FUNCTION "ROLL_PB2" : Void
{ S7_Optimized_Access := 'TRUE' }
VERSION : 0.1
VAR_TEMP
    r : Bool;
    a1 : Word;
    a2 : Word;
    activeDataBlock : Int;
    comparisonResults : Array[0..0] of Bool;
END_VAR
BEGIN
    #r := FALSE;
    #a1 := W#16#0000;
    #a2 := W#16#0000;
    #activeDataBlock := 0;
    // PB2, STEP 5 network 1
    #r := ((NOT "ROLL_State".M[0, 1]) AND "ROLL_State".S5Timers[11].Q);
    "ROLL_State".M[4, 1] := #r;
    // PB2, STEP 5 network 2
    #r := ((NOT "ROLL_State".M[4, 1]) OR "ROLL_IO".Input[1, 0]);
    "ROLL_State".M[3, 1] := #r;
    // PB2, STEP 5 network 3
    #r := ((((NOT "ROLL_State".M[31, 4]) AND "ROLL_IO".Input[0, 4] AND "ROLL_State".M[4, 1]) OR "ROLL_State".M[31, 5]) AND "ROLL_IO".Input[0, 2]);
    "ROLL_State".M[4, 4] := #r;
    // PB2, STEP 5 network 4
    #r := (NOT "ROLL_IO".Input[11, 7]);
    IF #r THEN "ROLL_State".M[5, 0] := TRUE; END_IF;
    #r := "ROLL_State".M[3, 1];
    IF #r THEN "ROLL_State".M[5, 0] := FALSE; END_IF;
    // PB2, STEP 5 network 5
    #r := (NOT "ROLL_IO".Input[13, 5]);
    IF #r THEN "ROLL_State".M[5, 1] := TRUE; END_IF;
    #r := "ROLL_State".M[3, 1];
    IF #r THEN "ROLL_State".M[5, 1] := FALSE; END_IF;
    // PB2, STEP 5 network 6
    #r := (NOT "ROLL_IO".Input[13, 0]);
    IF #r THEN "ROLL_State".M[5, 2] := TRUE; END_IF;
    #r := "ROLL_State".M[3, 1];
    IF #r THEN "ROLL_State".M[5, 2] := FALSE; END_IF;
    // PB2, STEP 5 network 7
    #r := (NOT "ROLL_IO".Input[8, 5]);
    IF #r THEN "ROLL_State".M[5, 3] := TRUE; END_IF;
    #r := "ROLL_State".M[3, 1];
    IF #r THEN "ROLL_State".M[5, 3] := FALSE; END_IF;
    // PB2, STEP 5 network 8
    #r := "ROLL_State".M[0, 3];
    IF #r THEN "ROLL_State".M[5, 4] := TRUE; END_IF;
    #r := "ROLL_State".M[3, 1];
    IF #r THEN "ROLL_State".M[5, 4] := FALSE; END_IF;
    // PB2, STEP 5 network 9
    #r := "ROLL_State".M[0, 3];
    IF #r THEN "ROLL_State".M[5, 5] := TRUE; END_IF;
    #r := "ROLL_State".M[3, 1];
    IF #r THEN "ROLL_State".M[5, 5] := FALSE; END_IF;
    // PB2, STEP 5 network 10
    #r := "ROLL_IO".Input[3, 6];
    IF #r THEN "ROLL_State".M[5, 6] := TRUE; END_IF;
    #r := "ROLL_State".M[3, 1];
    IF #r THEN "ROLL_State".M[5, 6] := FALSE; END_IF;
    // PB2, STEP 5 network 11
    #r := (NOT "ROLL_IO".Input[3, 7]);
    IF #r THEN "ROLL_State".M[5, 7] := TRUE; END_IF;
    #r := "ROLL_State".M[3, 1];
    IF #r THEN "ROLL_State".M[5, 7] := FALSE; END_IF;
    // PB2, STEP 5 network 12
    #r := (NOT "ROLL_IO".Input[5, 2]);
    IF #r THEN "ROLL_State".M[6, 0] := TRUE; END_IF;
    #r := ("ROLL_IO".Input[5, 2] AND "ROLL_State".M[3, 1]);
    IF #r THEN "ROLL_State".M[6, 0] := FALSE; END_IF;
    // PB2, STEP 5 network 13
    #r := ((NOT "ROLL_IO".Input[5, 3]) AND "ROLL_State".S5Timers[31].Q);
    IF #r THEN "ROLL_State".M[6, 1] := TRUE; END_IF;
    #r := "ROLL_State".M[3, 1];
    IF #r THEN "ROLL_State".M[6, 1] := FALSE; END_IF;
    // PB2, STEP 5 network 14
    #r := (NOT "ROLL_IO".Input[5, 4]);
    IF #r THEN "ROLL_State".M[6, 2] := TRUE; END_IF;
    #r := ("ROLL_IO".Input[5, 4] AND "ROLL_State".M[3, 1]);
    IF #r THEN "ROLL_State".M[6, 2] := FALSE; END_IF;
    // PB2, STEP 5 network 15
    #r := ((NOT "ROLL_IO".Input[5, 5]) AND "ROLL_State".M[40, 5] AND "ROLL_State".S5Timers[17].Q);
    IF #r THEN "ROLL_State".M[6, 3] := TRUE; END_IF;
    #r := "ROLL_State".M[3, 1];
    IF #r THEN "ROLL_State".M[6, 3] := FALSE; END_IF;
    // PB2, STEP 5 network 16
    #r := ((NOT "ROLL_IO".Input[6, 0]) AND "ROLL_State".S5Timers[32].Q);
    IF #r THEN "ROLL_State".M[6, 4] := TRUE; END_IF;
    #r := "ROLL_State".M[3, 1];
    IF #r THEN "ROLL_State".M[6, 4] := FALSE; END_IF;
    // PB2, STEP 5 network 17
    #r := ((NOT "ROLL_IO".Input[6, 2]) AND "ROLL_State".S5Timers[33].Q);
    IF #r THEN "ROLL_State".M[6, 5] := TRUE; END_IF;
    #r := "ROLL_State".M[3, 1];
    IF #r THEN "ROLL_State".M[6, 5] := FALSE; END_IF;
    // PB2, STEP 5 network 18
    #r := "ROLL_State".M[0, 3];
    IF #r THEN "ROLL_State".M[6, 6] := TRUE; END_IF;
    #r := "ROLL_State".M[3, 1];
    IF #r THEN "ROLL_State".M[6, 6] := FALSE; END_IF;
    // PB2, STEP 5 network 19
    #r := ((NOT "ROLL_State".M[0, 3]) AND "ROLL_State".S5Timers[35].Q);
    IF #r THEN "ROLL_State".M[6, 7] := TRUE; END_IF;
    #r := "ROLL_State".M[3, 1];
    IF #r THEN "ROLL_State".M[6, 7] := FALSE; END_IF;
    // PB2, STEP 5 network 20
    #r := ((NOT "ROLL_State".M[0, 3]) AND "ROLL_State".S5Timers[36].Q);
    IF #r THEN "ROLL_State".M[7, 0] := TRUE; END_IF;
    #r := "ROLL_State".M[3, 1];
    IF #r THEN "ROLL_State".M[7, 0] := FALSE; END_IF;
    // PB2, STEP 5 network 21
    #r := ((NOT "ROLL_State".M[0, 3]) AND "ROLL_State".M[48, 1] AND "ROLL_State".S5Timers[37].Q);
    IF #r THEN "ROLL_State".M[7, 1] := TRUE; END_IF;
    #r := "ROLL_State".M[3, 1];
    IF #r THEN "ROLL_State".M[7, 1] := FALSE; END_IF;
    // PB2, STEP 5 network 22
    #r := ((NOT "ROLL_State".M[0, 3]) AND "ROLL_State".S5Timers[38].Q);
    IF #r THEN "ROLL_State".M[7, 2] := TRUE; END_IF;
    #r := "ROLL_State".M[3, 1];
    IF #r THEN "ROLL_State".M[7, 2] := FALSE; END_IF;
    // PB2, STEP 5 network 23
    #r := ((NOT "ROLL_IO".Input[5, 6]) AND "ROLL_State".S5Timers[16].Q);
    IF #r THEN "ROLL_State".M[7, 3] := TRUE; END_IF;
    #r := ("ROLL_IO".Input[5, 6] AND "ROLL_State".M[3, 1]);
    IF #r THEN "ROLL_State".M[7, 3] := FALSE; END_IF;
    // PB2, STEP 5 network 24
    #r := "ROLL_State".M[0, 3];
    IF #r THEN "ROLL_State".M[7, 4] := TRUE; END_IF;
    #r := "ROLL_State".M[3, 1];
    IF #r THEN "ROLL_State".M[7, 4] := FALSE; END_IF;
    // PB2, STEP 5 network 25
    #r := "ROLL_State".M[0, 3];
    IF #r THEN "ROLL_State".M[7, 5] := TRUE; END_IF;
    #r := "ROLL_State".M[3, 1];
    IF #r THEN "ROLL_State".M[7, 5] := FALSE; END_IF;
    // PB2, STEP 5 network 26
    #r := "ROLL_State".M[0, 3];
    IF #r THEN "ROLL_State".M[7, 6] := TRUE; END_IF;
    #r := "ROLL_State".M[3, 1];
    IF #r THEN "ROLL_State".M[7, 6] := FALSE; END_IF;
    // PB2, STEP 5 network 27
    #r := (NOT "ROLL_IO".Input[6, 7]);
    IF #r THEN "ROLL_State".M[7, 7] := TRUE; END_IF;
    #r := "ROLL_State".M[3, 1];
    IF #r THEN "ROLL_State".M[7, 7] := FALSE; END_IF;
    // PB2, STEP 5 network 28
    #a2 := #a1;
    #a1 := W#16#1050;
    #r := ((NOT "ROLL_IO".Input[7, 6]) AND "ROLL_IO".Output[20, 5]);
    "ROLL_TimerOp"(Number := 30, Operation := 0, Signal := #r, Preset := #a1);
    #r := "ROLL_State".S5Timers[30].Q;
    IF #r THEN "ROLL_State".M[8, 6] := TRUE; END_IF;
    #r := "ROLL_State".M[3, 1];
    IF #r THEN "ROLL_State".M[8, 6] := FALSE; END_IF;
    // PB2, STEP 5 network 29
    #r := "ROLL_State".M[0, 3];
    IF #r THEN "ROLL_State".M[8, 7] := TRUE; END_IF;
    #r := "ROLL_State".M[3, 1];
    IF #r THEN "ROLL_State".M[8, 7] := FALSE; END_IF;
    // PB2, STEP 5 network 30
    #r := ((NOT "ROLL_IO".Input[13, 7]) AND "ROLL_State".M[4, 1]);
    IF #r THEN "ROLL_State".M[9, 0] := TRUE; END_IF;
    #r := ("ROLL_IO".Input[13, 7] AND "ROLL_State".M[3, 1]);
    IF #r THEN "ROLL_State".M[9, 0] := FALSE; END_IF;
    // PB2, STEP 5 network 31
    #r := "ROLL_State".M[0, 3];
    IF #r THEN "ROLL_State".M[9, 1] := TRUE; END_IF;
    #r := "ROLL_State".M[3, 1];
    IF #r THEN "ROLL_State".M[9, 1] := FALSE; END_IF;
    // PB2, STEP 5 network 32
    #r := ((NOT "ROLL_State".M[28, 4]) AND (NOT "ROLL_State".M[31, 5]) AND (((NOT "ROLL_State".M[20, 2]) AND ("ROLL_IO".Input[123, 5] OR "ROLL_IO".Input[123, 6])) OR "ROLL_State".M[70, 2] OR "ROLL_State".M[70, 3]) AND "ROLL_IO".Input[0, 4] AND "ROLL_State".M[4, 1]);
    IF #r THEN "ROLL_State".M[9, 2] := TRUE; END_IF;
    #r := "ROLL_State".M[3, 1];
    IF #r THEN "ROLL_State".M[9, 2] := FALSE; END_IF;
    // PB2, STEP 5 network 33
    #r := ("ROLL_State".M[4, 1] AND "ROLL_State".S5Timers[19].Q);
    IF #r THEN "ROLL_State".M[9, 3] := TRUE; END_IF;
    #r := "ROLL_State".M[3, 1];
    IF #r THEN "ROLL_State".M[9, 3] := FALSE; END_IF;
    // PB2, STEP 5 network 34
    #r := (((("ROLL_State".M[20, 4] OR "ROLL_State".M[20, 5]) AND "ROLL_IO".Input[0, 1] AND "ROLL_State".M[190, 6]) OR "ROLL_State".M[31, 5]) AND "ROLL_State".S5Timers[95].Q);
    "ROLL_State".M[9, 4] := #r;
    // PB2, STEP 5 network 35
    #r := "ROLL_State".M[0, 3];
    IF #r THEN "ROLL_State".M[9, 5] := TRUE; END_IF;
    #r := "ROLL_State".M[3, 1];
    IF #r THEN "ROLL_State".M[9, 5] := FALSE; END_IF;
    // PB2, STEP 5 network 36
    #r := "ROLL_State".M[0, 3];
    IF #r THEN "ROLL_State".M[9, 6] := TRUE; END_IF;
    #r := "ROLL_State".M[3, 1];
    IF #r THEN "ROLL_State".M[9, 6] := FALSE; END_IF;
    // PB2, STEP 5 network 37
    #r := "ROLL_State".M[0, 3];
    IF #r THEN "ROLL_State".M[9, 7] := TRUE; END_IF;
    #r := "ROLL_State".M[3, 1];
    IF #r THEN "ROLL_State".M[9, 7] := FALSE; END_IF;
    // PB2, STEP 5 network 38
    #r := ((NOT "ROLL_IO".Input[12, 0]) AND "ROLL_State".M[4, 1]);
    IF #r THEN "ROLL_State".M[10, 0] := TRUE; END_IF;
    #r := (((((NOT "ROLL_State".S5Timers[11].Q) AND "ROLL_IO".Input[3, 0]) OR "ROLL_IO".Input[12, 5]) AND "ROLL_State".M[3, 1]) OR (NOT "ROLL_State".M[4, 1]) OR "ROLL_State".M[0, 7]);
    IF #r THEN "ROLL_State".M[10, 0] := FALSE; END_IF;
    // PB2, STEP 5 network 39
    #r := ((NOT "ROLL_IO".Input[12, 6]) AND "ROLL_State".M[4, 1]);
    IF #r THEN "ROLL_State".M[10, 1] := TRUE; END_IF;
    #r := (((((NOT "ROLL_State".S5Timers[11].Q) AND "ROLL_IO".Input[3, 0]) OR "ROLL_IO".Input[12, 1]) AND "ROLL_State".M[3, 1]) OR (NOT "ROLL_State".M[4, 1]) OR "ROLL_State".M[0, 7]);
    IF #r THEN "ROLL_State".M[10, 1] := FALSE; END_IF;
    // PB2, STEP 5 network 40
    #r := "ROLL_State".M[0, 3];
    IF #r THEN "ROLL_State".M[10, 2] := TRUE; END_IF;
    #r := "ROLL_State".M[3, 1];
    IF #r THEN "ROLL_State".M[10, 2] := FALSE; END_IF;
    // PB2, STEP 5 network 41
    #r := "ROLL_State".M[0, 3];
    IF #r THEN "ROLL_State".M[10, 3] := TRUE; END_IF;
    #r := "ROLL_State".M[3, 1];
    IF #r THEN "ROLL_State".M[10, 3] := FALSE; END_IF;
    // PB2, STEP 5 network 42
    #r := "ROLL_State".M[0, 3];
    IF #r THEN "ROLL_State".M[10, 4] := TRUE; END_IF;
    #r := "ROLL_State".M[3, 1];
    IF #r THEN "ROLL_State".M[10, 4] := FALSE; END_IF;
    // PB2, STEP 5 network 43
    #r := "ROLL_State".M[0, 3];
    IF #r THEN "ROLL_State".M[10, 5] := TRUE; END_IF;
    #r := "ROLL_State".M[3, 1];
    IF #r THEN "ROLL_State".M[10, 5] := FALSE; END_IF;
    // PB2, STEP 5 network 44
    #r := "ROLL_State".M[0, 3];
    IF #r THEN "ROLL_State".M[10, 6] := TRUE; END_IF;
    #r := "ROLL_State".M[3, 1];
    IF #r THEN "ROLL_State".M[10, 6] := FALSE; END_IF;
    // PB2, STEP 5 network 45
    #r := "ROLL_State".M[0, 3];
    IF #r THEN "ROLL_State".M[10, 7] := TRUE; END_IF;
    #r := "ROLL_State".M[3, 1];
    IF #r THEN "ROLL_State".M[10, 7] := FALSE; END_IF;
    // PB2, STEP 5 network 46
    #r := ("ROLL_State".M[4, 1] AND "ROLL_State".M[63, 2]);
    IF #r THEN "ROLL_State".M[11, 0] := TRUE; END_IF;
    #r := "ROLL_State".M[3, 1];
    IF #r THEN "ROLL_State".M[11, 0] := FALSE; END_IF;
    // PB2, STEP 5 network 47
    #r := ("ROLL_IO".Input[13, 3] AND "ROLL_State".M[4, 1] AND "ROLL_State".S5Timers[112].Q);
    IF #r THEN "ROLL_State".M[11, 1] := TRUE; END_IF;
    #r := "ROLL_State".M[3, 1];
    IF #r THEN "ROLL_State".M[11, 1] := FALSE; END_IF;
    // PB2, STEP 5 network 48
    #r := ((NOT "ROLL_IO".Input[13, 3]) AND "ROLL_State".M[4, 1] AND "ROLL_State".S5Timers[15].Q);
    IF #r THEN "ROLL_State".M[11, 2] := TRUE; END_IF;
    #r := "ROLL_State".M[3, 1];
    IF #r THEN "ROLL_State".M[11, 2] := FALSE; END_IF;
    // PB2, STEP 5 network 49
    #r := ("ROLL_State".M[4, 1] AND "ROLL_State".M[63, 3]);
    IF #r THEN "ROLL_State".M[11, 3] := TRUE; END_IF;
    #r := "ROLL_State".M[3, 1];
    IF #r THEN "ROLL_State".M[11, 3] := FALSE; END_IF;
    // PB2, STEP 5 network 50
    #r := ("ROLL_State".M[190, 6] AND "ROLL_State".M[23, 2] AND "ROLL_State".M[60, 3]);
    IF #r THEN "ROLL_State".M[11, 4] := TRUE; END_IF;
    #r := "ROLL_State".M[3, 1];
    IF #r THEN "ROLL_State".M[11, 4] := FALSE; END_IF;
    // PB2, STEP 5 network 51
    #r := "ROLL_State".M[0, 3];
    IF #r THEN "ROLL_State".M[11, 5] := TRUE; END_IF;
    #r := "ROLL_State".M[3, 1];
    IF #r THEN "ROLL_State".M[11, 5] := FALSE; END_IF;
    // PB2, STEP 5 network 52
    #r := "ROLL_State".M[0, 3];
    IF #r THEN "ROLL_State".M[11, 6] := TRUE; END_IF;
    #r := "ROLL_State".M[3, 1];
    IF #r THEN "ROLL_State".M[11, 6] := FALSE; END_IF;
    // PB2, STEP 5 network 53
    #r := "ROLL_State".M[0, 3];
    IF #r THEN "ROLL_State".M[11, 7] := TRUE; END_IF;
    #r := "ROLL_State".M[3, 1];
    IF #r THEN "ROLL_State".M[11, 7] := FALSE; END_IF;
    // PB2, STEP 5 network 54
    #r := (NOT "ROLL_IO".Input[8, 3]);
    IF #r THEN "ROLL_State".M[12, 0] := TRUE; END_IF;
    #r := "ROLL_State".M[3, 1];
    IF #r THEN "ROLL_State".M[12, 0] := FALSE; END_IF;
    // PB2, STEP 5 network 55
    #r := ((NOT "ROLL_IO".Input[0, 7]) AND (NOT "ROLL_IO".Input[1, 4]) AND "ROLL_State".M[4, 4]);
    IF #r THEN "ROLL_State".M[12, 1] := TRUE; END_IF;
    #r := "ROLL_State".M[3, 1];
    IF #r THEN "ROLL_State".M[12, 1] := FALSE; END_IF;
    // PB2, STEP 5 network 56
    #r := "ROLL_State".M[0, 3];
    IF #r THEN "ROLL_State".M[12, 2] := TRUE; END_IF;
    #r := "ROLL_State".M[3, 1];
    IF #r THEN "ROLL_State".M[12, 2] := FALSE; END_IF;
    // PB2, STEP 5 network 57
    #r := "ROLL_State".M[0, 3];
    IF #r THEN "ROLL_State".M[12, 3] := TRUE; END_IF;
    #r := "ROLL_State".M[3, 1];
    IF #r THEN "ROLL_State".M[12, 3] := FALSE; END_IF;
    // PB2, STEP 5 network 58
    #r := "ROLL_State".M[0, 3];
    IF #r THEN "ROLL_State".M[13, 0] := TRUE; END_IF;
    #r := "ROLL_State".M[3, 1];
    IF #r THEN "ROLL_State".M[13, 0] := FALSE; END_IF;
    // PB2, STEP 5 network 59
    #r := (NOT "ROLL_IO".Input[3, 2]);
    IF #r THEN "ROLL_State".M[13, 1] := TRUE; END_IF;
    #r := "ROLL_State".M[3, 1];
    IF #r THEN "ROLL_State".M[13, 1] := FALSE; END_IF;
    // PB2, STEP 5 network 60
    #r := ((NOT "ROLL_IO".Input[4, 7]) AND "ROLL_IO".Input[0, 1] AND "ROLL_State".M[190, 6] AND "ROLL_State".M[27, 4]);
    IF #r THEN "ROLL_State".M[13, 2] := TRUE; END_IF;
    #r := "ROLL_State".M[3, 1];
    IF #r THEN "ROLL_State".M[13, 2] := FALSE; END_IF;
    // PB2, STEP 5 network 61
    #r := (NOT "ROLL_IO".Input[5, 0]);
    IF #r THEN "ROLL_State".M[13, 3] := TRUE; END_IF;
    #r := ("ROLL_IO".Input[5, 0] AND "ROLL_State".M[3, 1]);
    IF #r THEN "ROLL_State".M[13, 3] := FALSE; END_IF;
    // PB2, STEP 5 network 62
    #r := (NOT "ROLL_IO".Input[10, 7]);
    IF #r THEN "ROLL_State".M[13, 4] := TRUE; END_IF;
    #r := ("ROLL_IO".Input[10, 7] AND "ROLL_State".M[3, 1]);
    IF #r THEN "ROLL_State".M[13, 4] := FALSE; END_IF;
    // PB2, STEP 5 network 63
    #r := (NOT "ROLL_IO".Input[4, 5]);
    IF #r THEN "ROLL_State".M[13, 7] := TRUE; END_IF;
    #r := "ROLL_State".M[3, 1];
    IF #r THEN "ROLL_State".M[13, 7] := FALSE; END_IF;
    // PB2, STEP 5 network 64
    #a2 := #a1;
    #a1 := W#16#2020;
    #r := (((NOT "ROLL_IO".Input[10, 0]) OR (NOT "ROLL_IO".Input[10, 1]) OR (NOT "ROLL_IO".Input[10, 2]) OR (NOT "ROLL_IO".Input[10, 3])) AND "ROLL_IO".Output[19, 1]);
    "ROLL_TimerOp"(Number := 50, Operation := 0, Signal := #r, Preset := #a1);
    // PB2, STEP 5 network 65
    #r := ((NOT "ROLL_IO".Input[10, 0]) AND "ROLL_State".S5Timers[50].Q);
    IF #r THEN "ROLL_State".M[14, 0] := TRUE; END_IF;
    #r := "ROLL_State".M[3, 1];
    IF #r THEN "ROLL_State".M[14, 0] := FALSE; END_IF;
    // PB2, STEP 5 network 66
    #r := ((NOT "ROLL_IO".Input[10, 1]) AND "ROLL_State".S5Timers[50].Q);
    IF #r THEN "ROLL_State".M[14, 1] := TRUE; END_IF;
    #r := "ROLL_State".M[3, 1];
    IF #r THEN "ROLL_State".M[14, 1] := FALSE; END_IF;
    // PB2, STEP 5 network 67
    #r := ((NOT "ROLL_IO".Input[10, 2]) AND "ROLL_State".S5Timers[50].Q);
    IF #r THEN "ROLL_State".M[14, 2] := TRUE; END_IF;
    #r := "ROLL_State".M[3, 1];
    IF #r THEN "ROLL_State".M[14, 2] := FALSE; END_IF;
    // PB2, STEP 5 network 68
    #r := ((NOT "ROLL_IO".Input[10, 3]) AND "ROLL_State".S5Timers[50].Q);
    IF #r THEN "ROLL_State".M[14, 3] := TRUE; END_IF;
    #r := "ROLL_State".M[3, 1];
    IF #r THEN "ROLL_State".M[14, 3] := FALSE; END_IF;
    // PB2, STEP 5 network 69
    #r := "ROLL_State".M[0, 3];
    IF #r THEN "ROLL_State".M[15, 2] := TRUE; END_IF;
    #r := "ROLL_State".M[3, 1];
    IF #r THEN "ROLL_State".M[15, 2] := FALSE; END_IF;
    // PB2, STEP 5 network 70
    #r := "ROLL_State".M[0, 3];
    IF #r THEN "ROLL_State".M[15, 3] := TRUE; END_IF;
    #r := "ROLL_State".M[3, 1];
    IF #r THEN "ROLL_State".M[15, 3] := FALSE; END_IF;
    // PB2, STEP 5 network 71
    #r := "ROLL_State".M[0, 3];
    IF #r THEN "ROLL_State".M[15, 4] := TRUE; END_IF;
    #r := "ROLL_State".M[3, 1];
    IF #r THEN "ROLL_State".M[15, 4] := FALSE; END_IF;
    // PB2, STEP 5 network 72
    #r := (NOT "ROLL_IO".Input[4, 0]);
    IF #r THEN "ROLL_State".M[15, 5] := TRUE; END_IF;
    #r := "ROLL_State".M[3, 1];
    IF #r THEN "ROLL_State".M[15, 5] := FALSE; END_IF;
    // PB2, STEP 5 network 73
    #r := (NOT "ROLL_IO".Input[4, 1]);
    IF #r THEN "ROLL_State".M[15, 6] := TRUE; END_IF;
    #r := "ROLL_State".M[3, 1];
    IF #r THEN "ROLL_State".M[15, 6] := FALSE; END_IF;
    // PB2, STEP 5 network 74
    #r := (NOT "ROLL_IO".Input[4, 2]);
    IF #r THEN "ROLL_State".M[15, 7] := TRUE; END_IF;
    #r := "ROLL_State".M[3, 1];
    IF #r THEN "ROLL_State".M[15, 7] := FALSE; END_IF;
    // PB2, STEP 5 network 75
    #r := "ROLL_State".M[16, 0];
    IF #r THEN "ROLL_State".M[16, 0] := TRUE; END_IF;
    #r := "ROLL_State".M[3, 1];
    IF #r THEN "ROLL_State".M[16, 0] := FALSE; END_IF;
    // PB2, STEP 5 network 76
    #r := "ROLL_State".M[16, 1];
    IF #r THEN "ROLL_State".M[16, 1] := TRUE; END_IF;
    #r := "ROLL_State".M[3, 1];
    IF #r THEN "ROLL_State".M[16, 1] := FALSE; END_IF;
    // PB2, STEP 5 network 77
    #r := "ROLL_State".M[16, 2];
    IF #r THEN "ROLL_State".M[16, 2] := TRUE; END_IF;
    #r := "ROLL_State".M[3, 1];
    IF #r THEN "ROLL_State".M[16, 2] := FALSE; END_IF;
    // PB2, STEP 5 network 78
    #r := ("ROLL_State".M[34, 1] AND "ROLL_State".M[4, 1]);
    IF #r THEN "ROLL_State".M[16, 3] := TRUE; END_IF;
    #r := "ROLL_State".M[3, 1];
    IF #r THEN "ROLL_State".M[16, 3] := FALSE; END_IF;
    // PB2, STEP 5 network 79
    #r := "ROLL_State".M[16, 4];
    IF #r THEN "ROLL_State".M[16, 4] := TRUE; END_IF;
    #r := ((NOT "ROLL_IO".Input[123, 1]) AND (NOT "ROLL_IO".Input[123, 4]) AND (NOT "ROLL_IO".Input[123, 5]) AND (NOT "ROLL_IO".Input[123, 6]) AND (NOT "ROLL_IO".Input[125, 0]) AND (NOT "ROLL_IO".Input[125, 1]) AND "ROLL_State".M[3, 1]);
    IF #r THEN "ROLL_State".M[16, 4] := FALSE; END_IF;
    // PB2, STEP 5 network 80
    #r := "ROLL_State".M[16, 5];
    IF #r THEN "ROLL_State".M[16, 5] := TRUE; END_IF;
    #r := "ROLL_State".M[3, 1];
    IF #r THEN "ROLL_State".M[16, 5] := FALSE; END_IF;
    // PB2, STEP 5 network 81
    #r := ((NOT "ROLL_IO".Input[3, 4]) AND "ROLL_State".M[4, 1]);
    IF #r THEN "ROLL_State".M[16, 6] := TRUE; END_IF;
    #r := ("ROLL_IO".Input[3, 4] AND "ROLL_State".M[3, 1]);
    IF #r THEN "ROLL_State".M[16, 6] := FALSE; END_IF;
    // PB2, STEP 5 network 82
    #r := ((NOT "ROLL_IO".Input[3, 1]) AND ((("ROLL_State".M[190, 5] OR "ROLL_State".M[190, 6]) AND "ROLL_IO".Input[0, 1]) OR "ROLL_State".M[4, 4]) AND "ROLL_State".M[4, 1]);
    IF #r THEN "ROLL_State".M[16, 7] := TRUE; END_IF;
    #r := "ROLL_State".M[3, 1];
    IF #r THEN "ROLL_State".M[16, 7] := FALSE; END_IF;
    // PB2, STEP 5 network 83
    #r := ((NOT "ROLL_IO".Input[3, 5]) AND "ROLL_State".M[4, 1]);
    IF #r THEN "ROLL_State".M[17, 0] := TRUE; END_IF;
    #r := ("ROLL_IO".Input[3, 5] AND "ROLL_State".M[3, 1]);
    IF #r THEN "ROLL_State".M[17, 0] := FALSE; END_IF;
    // PB2, STEP 5 network 84
    #r := "ROLL_State".M[0, 3];
    IF #r THEN "ROLL_State".M[17, 1] := TRUE; END_IF;
    #r := "ROLL_State".M[3, 1];
    IF #r THEN "ROLL_State".M[17, 1] := FALSE; END_IF;
    // PB2, STEP 5 network 85
    #r := "ROLL_State".M[0, 3];
    IF #r THEN "ROLL_State".M[17, 2] := TRUE; END_IF;
    #r := "ROLL_State".M[3, 1];
    IF #r THEN "ROLL_State".M[17, 2] := FALSE; END_IF;
    // PB2, STEP 5 network 86
    #r := "ROLL_State".M[0, 3];
    IF #r THEN "ROLL_State".M[17, 3] := TRUE; END_IF;
    #r := "ROLL_State".M[3, 1];
    IF #r THEN "ROLL_State".M[17, 3] := FALSE; END_IF;
    // PB2, STEP 5 network 87
    #r := "ROLL_State".M[0, 3];
    IF #r THEN "ROLL_State".M[17, 4] := TRUE; END_IF;
    #r := "ROLL_State".M[3, 1];
    IF #r THEN "ROLL_State".M[17, 4] := FALSE; END_IF;
    // PB2, STEP 5 network 88
    #r := "ROLL_State".M[0, 3];
    IF #r THEN "ROLL_State".M[17, 5] := TRUE; END_IF;
    #r := "ROLL_State".M[3, 1];
    IF #r THEN "ROLL_State".M[17, 5] := FALSE; END_IF;
    // PB2, STEP 5 network 89
    #r := "ROLL_State".M[0, 3];
    IF #r THEN "ROLL_State".M[17, 6] := TRUE; END_IF;
    #r := "ROLL_State".M[3, 1];
    IF #r THEN "ROLL_State".M[17, 6] := FALSE; END_IF;
    // PB2, STEP 5 network 90
    #r := "ROLL_State".M[0, 3];
    IF #r THEN "ROLL_State".M[17, 7] := TRUE; END_IF;
    #r := "ROLL_State".M[3, 1];
    IF #r THEN "ROLL_State".M[17, 7] := FALSE; END_IF;
    // PB2, STEP 5 network 91
    #r := "ROLL_State".M[0, 3];
    IF #r THEN "ROLL_State".M[18, 0] := TRUE; END_IF;
    #r := "ROLL_State".M[3, 1];
    IF #r THEN "ROLL_State".M[18, 0] := FALSE; END_IF;
    // PB2, STEP 5 network 92
    #r := ((NOT "ROLL_IO".Input[14, 0]) AND ((("ROLL_State".M[190, 5] OR "ROLL_State".M[190, 6]) AND ("ROLL_State".M[23, 0] OR "ROLL_State".M[23, 1] OR "ROLL_State".M[23, 2] OR "ROLL_State".M[23, 3])) OR ("ROLL_State".M[16, 3] AND "ROLL_State".M[31, 4] AND "ROLL_State".M[37, 2]) OR "ROLL_State".M[74, 0]));
    IF #r THEN "ROLL_State".M[18, 1] := TRUE; END_IF;
    #r := "ROLL_State".M[3, 1];
    IF #r THEN "ROLL_State".M[18, 1] := FALSE; END_IF;
    // PB2, STEP 5 network 93
    #r := "ROLL_State".M[0, 3];
    IF #r THEN "ROLL_State".M[18, 2] := TRUE; END_IF;
    #r := "ROLL_State".M[3, 1];
    IF #r THEN "ROLL_State".M[18, 2] := FALSE; END_IF;
    // PB2, STEP 5 network 94
    #r := "ROLL_State".M[0, 3];
    IF #r THEN "ROLL_State".M[18, 3] := TRUE; END_IF;
    #r := "ROLL_State".M[3, 1];
    IF #r THEN "ROLL_State".M[18, 3] := FALSE; END_IF;
    // PB2, STEP 5 network 95
    #r := "ROLL_State".M[0, 3];
    IF #r THEN "ROLL_State".M[18, 4] := TRUE; END_IF;
    #r := "ROLL_State".M[3, 1];
    IF #r THEN "ROLL_State".M[18, 4] := FALSE; END_IF;
    // PB2, STEP 5 network 96
    #r := "ROLL_State".M[0, 3];
    IF #r THEN "ROLL_State".M[18, 5] := TRUE; END_IF;
    #r := "ROLL_State".M[3, 1];
    IF #r THEN "ROLL_State".M[18, 5] := FALSE; END_IF;
    // PB2, STEP 5 network 97
    #r := "ROLL_State".M[0, 3];
    IF #r THEN "ROLL_State".M[18, 6] := TRUE; END_IF;
    #r := "ROLL_State".M[3, 1];
    IF #r THEN "ROLL_State".M[18, 6] := FALSE; END_IF;
    // PB2, STEP 5 network 98
    #r := "ROLL_State".M[0, 3];
    IF #r THEN "ROLL_State".M[18, 7] := TRUE; END_IF;
    #r := "ROLL_State".M[3, 1];
    IF #r THEN "ROLL_State".M[18, 7] := FALSE; END_IF;
    // PB2, STEP 5 network 99
    #r := "ROLL_State".M[0, 3];
    IF #r THEN "ROLL_State".M[19, 0] := TRUE; END_IF;
    #r := "ROLL_State".M[3, 1];
    IF #r THEN "ROLL_State".M[19, 0] := FALSE; END_IF;
    // PB2, STEP 5 network 100
    #r := "ROLL_State".M[0, 3];
    IF #r THEN "ROLL_State".M[19, 1] := TRUE; END_IF;
    #r := "ROLL_State".M[3, 1];
    IF #r THEN "ROLL_State".M[19, 1] := FALSE; END_IF;
    // PB2, STEP 5 network 101
    #r := "ROLL_State".M[0, 3];
    IF #r THEN "ROLL_State".M[19, 2] := TRUE; END_IF;
    #r := "ROLL_State".M[3, 1];
    IF #r THEN "ROLL_State".M[19, 2] := FALSE; END_IF;
    // PB2, STEP 5 network 102
    #r := "ROLL_State".M[0, 3];
    IF #r THEN "ROLL_State".M[19, 3] := TRUE; END_IF;
    #r := "ROLL_State".M[3, 1];
    IF #r THEN "ROLL_State".M[19, 3] := FALSE; END_IF;
    // PB2, STEP 5 network 103
    #r := "ROLL_State".M[0, 3];
    IF #r THEN "ROLL_State".M[19, 4] := TRUE; END_IF;
    #r := "ROLL_State".M[3, 1];
    IF #r THEN "ROLL_State".M[19, 4] := FALSE; END_IF;
    // PB2, STEP 5 network 104
    #r := "ROLL_State".M[0, 3];
    IF #r THEN "ROLL_State".M[19, 5] := TRUE; END_IF;
    #r := "ROLL_State".M[3, 1];
    IF #r THEN "ROLL_State".M[19, 5] := FALSE; END_IF;
    // PB2, STEP 5 network 105
    #r := "ROLL_State".M[0, 3];
    IF #r THEN "ROLL_State".M[19, 6] := TRUE; END_IF;
    #r := "ROLL_State".M[3, 1];
    IF #r THEN "ROLL_State".M[19, 6] := FALSE; END_IF;
    // PB2, STEP 5 network 106
    #r := "ROLL_State".M[0, 3];
    IF #r THEN "ROLL_State".M[19, 7] := TRUE; END_IF;
    #r := "ROLL_State".M[3, 1];
    IF #r THEN "ROLL_State".M[19, 7] := FALSE; END_IF;
    // PB2, STEP 5 network 107
    RETURN;
END_FUNCTION

FUNCTION "ROLL_PB3" : Void
{ S7_Optimized_Access := 'TRUE' }
VERSION : 0.1
VAR_TEMP
    r : Bool;
    a1 : Word;
    a2 : Word;
    activeDataBlock : Int;
    comparisonResults : Array[0..15] of Bool;
END_VAR
BEGIN
    #r := FALSE;
    #a1 := W#16#0000;
    #a2 := W#16#0000;
    #activeDataBlock := 0;
    // PB3, STEP 5 network 1
    #a2 := #a1;
    #a1 := "ROLL_GetM"(FirstByte := 239, Width := 8);
    #a2 := #a1;
    #a1 := W#16#0001;
    #comparisonResults[0] := (WORD_TO_INT(#a2) = WORD_TO_INT(#a1));
    #r := #comparisonResults[0];
    "ROLL_State".M[20, 1] := #r;
    // PB3, STEP 5 network 2
    #a2 := #a1;
    #a1 := "ROLL_GetM"(FirstByte := 239, Width := 8);
    #a2 := #a1;
    #a1 := W#16#0002;
    #comparisonResults[1] := (WORD_TO_INT(#a2) = WORD_TO_INT(#a1));
    #r := #comparisonResults[1];
    "ROLL_State".M[20, 2] := #r;
    // PB3, STEP 5 network 3
    #a2 := #a1;
    #a1 := "ROLL_GetM"(FirstByte := 239, Width := 8);
    #a2 := #a1;
    #a1 := W#16#0003;
    #comparisonResults[2] := (WORD_TO_INT(#a2) = WORD_TO_INT(#a1));
    #r := #comparisonResults[2];
    "ROLL_State".M[20, 3] := #r;
    // PB3, STEP 5 network 4
    #a2 := #a1;
    #a1 := "ROLL_GetM"(FirstByte := 239, Width := 8);
    #a2 := #a1;
    #a1 := W#16#0004;
    #comparisonResults[3] := (WORD_TO_INT(#a2) = WORD_TO_INT(#a1));
    #r := #comparisonResults[3];
    "ROLL_State".M[20, 4] := #r;
    // PB3, STEP 5 network 5
    #a2 := #a1;
    #a1 := "ROLL_GetM"(FirstByte := 239, Width := 8);
    #a2 := #a1;
    #a1 := W#16#0005;
    #comparisonResults[4] := (WORD_TO_INT(#a2) = WORD_TO_INT(#a1));
    #r := #comparisonResults[4];
    "ROLL_State".M[20, 5] := #r;
    // PB3, STEP 5 network 6
    #a2 := #a1;
    #a1 := "ROLL_GetM"(FirstByte := 239, Width := 8);
    #a2 := #a1;
    #a1 := W#16#0007;
    #comparisonResults[5] := (WORD_TO_INT(#a2) = WORD_TO_INT(#a1));
    #r := #comparisonResults[5];
    "ROLL_State".M[20, 7] := #r;
    // PB3, STEP 5 network 7
    #a2 := #a1;
    #a1 := "ROLL_GetM"(FirstByte := 239, Width := 8);
    #a2 := #a1;
    #a1 := W#16#000A;
    #comparisonResults[6] := (WORD_TO_INT(#a2) = WORD_TO_INT(#a1));
    #r := #comparisonResults[6];
    "ROLL_State".M[22, 0] := #r;
    // PB3, STEP 5 network 8
    #a2 := #a1;
    #a1 := "ROLL_GetM"(FirstByte := 239, Width := 8);
    #a2 := #a1;
    #a1 := W#16#000B;
    #comparisonResults[7] := (WORD_TO_INT(#a2) = WORD_TO_INT(#a1));
    #r := #comparisonResults[7];
    "ROLL_State".M[22, 1] := #r;
    // PB3, STEP 5 network 9
    #a2 := #a1;
    #a1 := "ROLL_GetM"(FirstByte := 239, Width := 8);
    #a2 := #a1;
    #a1 := W#16#000C;
    #comparisonResults[8] := (WORD_TO_INT(#a2) = WORD_TO_INT(#a1));
    #r := #comparisonResults[8];
    "ROLL_State".M[22, 2] := #r;
    // PB3, STEP 5 network 10
    #a2 := #a1;
    #a1 := "ROLL_GetM"(FirstByte := 239, Width := 8);
    #a2 := #a1;
    #a1 := W#16#000D;
    #comparisonResults[9] := (WORD_TO_INT(#a2) = WORD_TO_INT(#a1));
    #r := #comparisonResults[9];
    "ROLL_State".M[22, 3] := #r;
    // PB3, STEP 5 network 11
    #a2 := #a1;
    #a1 := "ROLL_GetM"(FirstByte := 239, Width := 8);
    #a2 := #a1;
    #a1 := W#16#000E;
    #comparisonResults[10] := (WORD_TO_INT(#a2) = WORD_TO_INT(#a1));
    #r := #comparisonResults[10];
    "ROLL_State".M[22, 4] := #r;
    // PB3, STEP 5 network 12
    #a2 := #a1;
    #a1 := "ROLL_GetM"(FirstByte := 239, Width := 8);
    #a2 := #a1;
    #a1 := W#16#000F;
    #comparisonResults[11] := (WORD_TO_INT(#a2) = WORD_TO_INT(#a1));
    #r := #comparisonResults[11];
    "ROLL_State".M[22, 5] := #r;
    // PB3, STEP 5 network 13
    #a2 := #a1;
    #a1 := "ROLL_GetM"(FirstByte := 239, Width := 8);
    #a2 := #a1;
    #a1 := W#16#0014;
    #comparisonResults[12] := (WORD_TO_INT(#a2) = WORD_TO_INT(#a1));
    #r := #comparisonResults[12];
    "ROLL_State".M[23, 0] := #r;
    // PB3, STEP 5 network 14
    #a2 := #a1;
    #a1 := "ROLL_GetM"(FirstByte := 239, Width := 8);
    #a2 := #a1;
    #a1 := W#16#0015;
    #comparisonResults[13] := (WORD_TO_INT(#a2) = WORD_TO_INT(#a1));
    #r := #comparisonResults[13];
    "ROLL_State".M[23, 1] := #r;
    // PB3, STEP 5 network 15
    #a2 := #a1;
    #a1 := "ROLL_GetM"(FirstByte := 239, Width := 8);
    #a2 := #a1;
    #a1 := W#16#0016;
    #comparisonResults[14] := (WORD_TO_INT(#a2) = WORD_TO_INT(#a1));
    #r := #comparisonResults[14];
    "ROLL_State".M[23, 2] := #r;
    // PB3, STEP 5 network 16
    #a2 := #a1;
    #a1 := "ROLL_GetM"(FirstByte := 239, Width := 8);
    #a2 := #a1;
    #a1 := W#16#0017;
    #comparisonResults[15] := (WORD_TO_INT(#a2) = WORD_TO_INT(#a1));
    #r := #comparisonResults[15];
    "ROLL_State".M[23, 3] := #r;
    // PB3, STEP 5 network 17
    RETURN;
END_FUNCTION

FUNCTION "ROLL_PB4" : Void
{ S7_Optimized_Access := 'TRUE' }
VERSION : 0.1
VAR_TEMP
    r : Bool;
    a1 : Word;
    a2 : Word;
    activeDataBlock : Int;
    comparisonResults : Array[0..24] of Bool;
END_VAR
BEGIN
    #r := FALSE;
    #a1 := W#16#0000;
    #a2 := W#16#0000;
    #activeDataBlock := 0;
    // PB4, STEP 5 network 1
    #a2 := #a1;
    #a1 := "ROLL_GetM"(FirstByte := 239, Width := 8);
    #a2 := #a1;
    #a1 := W#16#001E;
    #comparisonResults[0] := (WORD_TO_INT(#a2) = WORD_TO_INT(#a1));
    #r := #comparisonResults[0];
    "ROLL_State".M[23, 5] := #r;
    // PB4, STEP 5 network 2
    #a2 := #a1;
    #a1 := "ROLL_GetM"(FirstByte := 239, Width := 8);
    #a2 := #a1;
    #a1 := W#16#001F;
    #comparisonResults[1] := (WORD_TO_INT(#a2) = WORD_TO_INT(#a1));
    #r := #comparisonResults[1];
    "ROLL_State".M[23, 6] := #r;
    // PB4, STEP 5 network 3
    #a2 := #a1;
    #a1 := "ROLL_GetM"(FirstByte := 239, Width := 8);
    #a2 := #a1;
    #a1 := W#16#0023;
    #comparisonResults[2] := (WORD_TO_INT(#a2) = WORD_TO_INT(#a1));
    #r := #comparisonResults[2];
    "ROLL_State".M[24, 0] := #r;
    // PB4, STEP 5 network 4
    #a2 := #a1;
    #a1 := "ROLL_GetM"(FirstByte := 239, Width := 8);
    #a2 := #a1;
    #a1 := W#16#0024;
    #comparisonResults[3] := (WORD_TO_INT(#a2) = WORD_TO_INT(#a1));
    #r := #comparisonResults[3];
    "ROLL_State".M[24, 1] := #r;
    // PB4, STEP 5 network 5
    #a2 := #a1;
    #a1 := "ROLL_GetM"(FirstByte := 239, Width := 8);
    #a2 := #a1;
    #a1 := W#16#0025;
    #comparisonResults[4] := (WORD_TO_INT(#a2) = WORD_TO_INT(#a1));
    #r := #comparisonResults[4];
    "ROLL_State".M[24, 2] := #r;
    // PB4, STEP 5 network 6
    #a2 := #a1;
    #a1 := "ROLL_GetM"(FirstByte := 239, Width := 8);
    #a2 := #a1;
    #a1 := W#16#0026;
    #comparisonResults[5] := (WORD_TO_INT(#a2) = WORD_TO_INT(#a1));
    #r := #comparisonResults[5];
    "ROLL_State".M[24, 3] := #r;
    // PB4, STEP 5 network 7
    #a2 := #a1;
    #a1 := "ROLL_GetM"(FirstByte := 239, Width := 8);
    #a2 := #a1;
    #a1 := W#16#0027;
    #comparisonResults[6] := (WORD_TO_INT(#a2) = WORD_TO_INT(#a1));
    #r := #comparisonResults[6];
    "ROLL_State".M[24, 4] := #r;
    // PB4, STEP 5 network 8
    #a2 := #a1;
    #a1 := "ROLL_GetM"(FirstByte := 239, Width := 8);
    #a2 := #a1;
    #a1 := W#16#0032;
    #comparisonResults[7] := (WORD_TO_INT(#a2) = WORD_TO_INT(#a1));
    #r := #comparisonResults[7];
    "ROLL_State".M[25, 0] := #r;
    // PB4, STEP 5 network 9
    #a2 := #a1;
    #a1 := "ROLL_GetM"(FirstByte := 239, Width := 8);
    #a2 := #a1;
    #a1 := W#16#0033;
    #comparisonResults[8] := (WORD_TO_INT(#a2) = WORD_TO_INT(#a1));
    #r := #comparisonResults[8];
    "ROLL_State".M[25, 1] := #r;
    // PB4, STEP 5 network 10
    #a2 := #a1;
    #a1 := "ROLL_GetM"(FirstByte := 239, Width := 8);
    #a2 := #a1;
    #a1 := W#16#0034;
    #comparisonResults[9] := (WORD_TO_INT(#a2) = WORD_TO_INT(#a1));
    #r := #comparisonResults[9];
    "ROLL_State".M[25, 2] := #r;
    // PB4, STEP 5 network 11
    #a2 := #a1;
    #a1 := "ROLL_GetM"(FirstByte := 239, Width := 8);
    #a2 := #a1;
    #a1 := W#16#0035;
    #comparisonResults[10] := (WORD_TO_INT(#a2) = WORD_TO_INT(#a1));
    #r := #comparisonResults[10];
    "ROLL_State".M[25, 3] := #r;
    // PB4, STEP 5 network 12
    #a2 := #a1;
    #a1 := "ROLL_GetM"(FirstByte := 239, Width := 8);
    #a2 := #a1;
    #a1 := W#16#0037;
    #comparisonResults[11] := (WORD_TO_INT(#a2) = WORD_TO_INT(#a1));
    #r := #comparisonResults[11];
    "ROLL_State".M[25, 4] := #r;
    // PB4, STEP 5 network 13
    #a2 := #a1;
    #a1 := "ROLL_GetM"(FirstByte := 239, Width := 8);
    #a2 := #a1;
    #a1 := W#16#0038;
    #comparisonResults[12] := (WORD_TO_INT(#a2) = WORD_TO_INT(#a1));
    #r := #comparisonResults[12];
    "ROLL_State".M[25, 5] := #r;
    // PB4, STEP 5 network 14
    #a2 := #a1;
    #a1 := "ROLL_GetM"(FirstByte := 239, Width := 8);
    #a2 := #a1;
    #a1 := W#16#0039;
    #comparisonResults[13] := (WORD_TO_INT(#a2) = WORD_TO_INT(#a1));
    #r := #comparisonResults[13];
    "ROLL_State".M[25, 6] := #r;
    // PB4, STEP 5 network 15
    #a2 := #a1;
    #a1 := "ROLL_GetM"(FirstByte := 239, Width := 8);
    #a2 := #a1;
    #a1 := W#16#003A;
    #comparisonResults[14] := (WORD_TO_INT(#a2) = WORD_TO_INT(#a1));
    #r := #comparisonResults[14];
    "ROLL_State".M[25, 7] := #r;
    // PB4, STEP 5 network 16
    #a2 := #a1;
    #a1 := "ROLL_GetM"(FirstByte := 239, Width := 8);
    #a2 := #a1;
    #a1 := W#16#003C;
    #comparisonResults[15] := (WORD_TO_INT(#a2) = WORD_TO_INT(#a1));
    #r := #comparisonResults[15];
    "ROLL_State".M[26, 0] := #r;
    // PB4, STEP 5 network 17
    #a2 := #a1;
    #a1 := "ROLL_GetM"(FirstByte := 239, Width := 8);
    #a2 := #a1;
    #a1 := W#16#003D;
    #comparisonResults[16] := (WORD_TO_INT(#a2) = WORD_TO_INT(#a1));
    #r := #comparisonResults[16];
    "ROLL_State".M[26, 1] := #r;
    // PB4, STEP 5 network 18
    #a2 := #a1;
    #a1 := "ROLL_GetM"(FirstByte := 239, Width := 8);
    #a2 := #a1;
    #a1 := W#16#003E;
    #comparisonResults[17] := (WORD_TO_INT(#a2) = WORD_TO_INT(#a1));
    #r := #comparisonResults[17];
    "ROLL_State".M[26, 2] := #r;
    // PB4, STEP 5 network 19
    #a2 := #a1;
    #a1 := "ROLL_GetM"(FirstByte := 239, Width := 8);
    #a2 := #a1;
    #a1 := W#16#003F;
    #comparisonResults[18] := (WORD_TO_INT(#a2) = WORD_TO_INT(#a1));
    #r := #comparisonResults[18];
    "ROLL_State".M[26, 3] := #r;
    // PB4, STEP 5 network 20
    #a2 := #a1;
    #a1 := "ROLL_GetM"(FirstByte := 239, Width := 8);
    #a2 := #a1;
    #a1 := W#16#0041;
    #comparisonResults[19] := (WORD_TO_INT(#a2) = WORD_TO_INT(#a1));
    #r := #comparisonResults[19];
    "ROLL_State".M[26, 5] := #r;
    // PB4, STEP 5 network 21
    #a2 := #a1;
    #a1 := "ROLL_GetM"(FirstByte := 239, Width := 8);
    #a2 := #a1;
    #a1 := W#16#0042;
    #comparisonResults[20] := (WORD_TO_INT(#a2) = WORD_TO_INT(#a1));
    #r := #comparisonResults[20];
    "ROLL_State".M[26, 6] := #r;
    // PB4, STEP 5 network 22
    #a2 := #a1;
    #a1 := "ROLL_GetM"(FirstByte := 239, Width := 8);
    #a2 := #a1;
    #a1 := W#16#0045;
    #comparisonResults[21] := (WORD_TO_INT(#a2) = WORD_TO_INT(#a1));
    #r := #comparisonResults[21];
    "ROLL_State".M[27, 1] := #r;
    // PB4, STEP 5 network 23
    #a2 := #a1;
    #a1 := "ROLL_GetM"(FirstByte := 239, Width := 8);
    #a2 := #a1;
    #a1 := W#16#0048;
    #comparisonResults[22] := (WORD_TO_INT(#a2) = WORD_TO_INT(#a1));
    #r := #comparisonResults[22];
    "ROLL_State".M[27, 4] := #r;
    // PB4, STEP 5 network 24
    #a2 := #a1;
    #a1 := "ROLL_GetM"(FirstByte := 239, Width := 8);
    #a2 := #a1;
    #a1 := W#16#0049;
    #comparisonResults[23] := (WORD_TO_INT(#a2) = WORD_TO_INT(#a1));
    #r := #comparisonResults[23];
    "ROLL_State".M[27, 5] := #r;
    // PB4, STEP 5 network 25
    #a2 := #a1;
    #a1 := "ROLL_GetM"(FirstByte := 239, Width := 8);
    #a2 := #a1;
    #a1 := W#16#0063;
    #comparisonResults[24] := (WORD_TO_INT(#a2) = WORD_TO_INT(#a1));
    #r := #comparisonResults[24];
    "ROLL_State".M[27, 7] := #r;
    // PB4, STEP 5 network 26
    RETURN;
END_FUNCTION

FUNCTION "ROLL_PB7" : Void
{ S7_Optimized_Access := 'TRUE' }
VERSION : 0.1
VAR_TEMP
    r : Bool;
    a1 : Word;
    a2 : Word;
    activeDataBlock : Int;
    comparisonResults : Array[0..0] of Bool;
END_VAR
BEGIN
    #r := FALSE;
    #a1 := W#16#0000;
    #a2 := W#16#0000;
    #activeDataBlock := 0;
    // PB7, STEP 5 network 1
    #r := ((NOT "ROLL_State".M[70, 2]) AND (NOT "ROLL_State".M[70, 3]) AND (NOT "ROLL_State".M[70, 4]) AND (NOT "ROLL_State".M[70, 6]) AND "ROLL_IO".Input[11, 0] AND "ROLL_IO".Input[11, 6] AND "ROLL_IO".Input[13, 3] AND "ROLL_State".M[63, 1]);
    "ROLL_State".M[28, 0] := #r;
    // PB7, STEP 5 network 2
    #r := ("ROLL_IO".Input[12, 1] AND "ROLL_IO".Input[12, 7]);
    "ROLL_State".M[28, 1] := #r;
    // PB7, STEP 5 network 3
    #r := ((NOT "ROLL_IO".Output[112, 5]) AND ((NOT "ROLL_IO".Output[112, 0]) OR (NOT "ROLL_State".M[31, 4])));
    "ROLL_State".M[28, 2] := #r;
    // PB7, STEP 5 network 4
    #r := (((NOT "ROLL_IO".Output[113, 0]) AND (NOT "ROLL_IO".Output[113, 1]) AND (NOT "ROLL_IO".Output[113, 3]) AND (NOT "ROLL_IO".Output[113, 5]) AND (NOT "ROLL_IO".Input[123, 5]) AND (NOT "ROLL_IO".Input[123, 6]) AND "ROLL_IO".Output[113, 2] AND "ROLL_IO".Output[113, 4] AND "ROLL_IO".Input[124, 1] AND "ROLL_IO".Input[124, 4]) OR "ROLL_State".M[0, 4]);
    "ROLL_State".M[240, 0] := #r;
    // PB7, STEP 5 network 5
    #r := ((((NOT "ROLL_IO".Output[113, 2]) AND "ROLL_IO".Output[113, 3] AND "ROLL_IO".Input[123, 5] AND "ROLL_IO".Input[124, 1] AND "ROLL_IO".Input[124, 4]) OR ((NOT "ROLL_IO".Output[113, 3]) AND "ROLL_IO".Output[113, 2] AND "ROLL_IO".Input[124, 1] AND "ROLL_IO".Input[124, 5]) OR "ROLL_State".M[0, 4]) AND "ROLL_State".M[20, 2]);
    "ROLL_State".M[240, 1] := #r;
    // PB7, STEP 5 network 6
    #r := ("ROLL_State".M[240, 0] OR "ROLL_State".M[240, 1]);
    "ROLL_State".M[28, 3] := #r;
    // PB7, STEP 5 network 7
    #r := ("ROLL_State".M[28, 0] AND "ROLL_State".M[28, 1] AND "ROLL_State".M[28, 2] AND "ROLL_State".M[28, 3]);
    "ROLL_State".M[28, 4] := #r;
    // PB7, STEP 5 network 8
    #r := ("ROLL_IO".Input[10, 7] AND "ROLL_IO".Input[3, 4] AND "ROLL_IO".Input[3, 5] AND "ROLL_IO".Input[3, 7]);
    "ROLL_State".M[28, 5] := #r;
    // PB7, STEP 5 network 9
    #r := ((NOT "ROLL_State".M[13, 4]) AND (NOT "ROLL_State".M[16, 6]) AND (NOT "ROLL_State".M[5, 7]) AND "ROLL_State".M[28, 5]);
    "ROLL_State".M[28, 6] := #r;
    // PB7, STEP 5 network 10
    #r := (("ROLL_IO".Input[0, 2] AND "ROLL_IO".Input[0, 4]) OR "ROLL_IO".Input[0, 1]);
    IF #r THEN "ROLL_State".M[29, 0] := TRUE; END_IF;
    #r := (NOT "ROLL_State".M[28, 6]);
    IF #r THEN "ROLL_State".M[29, 0] := FALSE; END_IF;
    // PB7, STEP 5 network 11
    #r := ("ROLL_State".M[29, 0] AND "ROLL_State".S5Timers[13].Q);
    "ROLL_State".M[29, 1] := #r;
    // PB7, STEP 5 network 12
    #r := (NOT "ROLL_State".M[12, 1]);
    "ROLL_State".M[30, 0] := #r;
    // PB7, STEP 5 network 13
    #r := "ROLL_State".M[0, 4];
    "ROLL_State".M[30, 1] := #r;
    // PB7, STEP 5 network 14
    #r := ((NOT "ROLL_State".M[6, 1]) AND (NOT "ROLL_State".M[6, 3]) AND (NOT "ROLL_State".M[6, 4]) AND (NOT "ROLL_State".M[6, 5]) AND (NOT "ROLL_State".M[6, 6]) AND (NOT "ROLL_State".M[6, 7]) AND (NOT "ROLL_State".M[7, 0]) AND (NOT "ROLL_State".M[7, 1]) AND (NOT "ROLL_State".M[7, 2]) AND (NOT "ROLL_State".M[7, 3]) AND (NOT "ROLL_State".M[7, 7]));
    "ROLL_State".M[30, 2] := #r;
    // PB7, STEP 5 network 15
    #r := ((NOT "ROLL_IO".Input[3, 6]) AND (NOT "ROLL_State".M[5, 6]));
    "ROLL_State".M[30, 3] := #r;
    // PB7, STEP 5 network 16
    #r := (("ROLL_State".M[30, 0] AND "ROLL_State".M[30, 1] AND "ROLL_State".M[30, 2] AND "ROLL_State".M[30, 3]) OR "ROLL_IO".Input[0, 0] OR "ROLL_IO".Input[0, 6]);
    "ROLL_State".M[30, 5] := #r;
    // PB7, STEP 5 network 17
    #r := ((NOT "ROLL_State".M[11, 0]) AND (NOT "ROLL_State".M[13, 1]) AND (NOT "ROLL_State".M[13, 3]) AND (NOT "ROLL_State".M[5, 0]) AND (NOT "ROLL_State".M[5, 1]) AND (NOT "ROLL_State".M[5, 2]));
    "ROLL_State".M[30, 6] := #r;
    // PB7, STEP 5 network 18
    #r := ((NOT "ROLL_State".M[11, 1]) AND (NOT "ROLL_State".M[5, 3]) AND (NOT "ROLL_State".M[9, 1]) AND (NOT "ROLL_State".M[9, 2]) AND (NOT "ROLL_State".M[9, 3]) AND "ROLL_IO".Input[8, 5] AND "ROLL_State".M[28, 6]);
    "ROLL_State".M[30, 7] := #r;
    // PB7, STEP 5 network 19
    #r := ((NOT "ROLL_State".M[12, 0]) AND (NOT "ROLL_State".M[9, 0]));
    "ROLL_State".M[31, 0] := #r;
    // PB7, STEP 5 network 20
    #r := ((NOT "ROLL_State".M[87, 5]) AND (NOT "ROLL_State".M[88, 1]) AND (NOT "ROLL_State".M[88, 3]) AND (NOT "ROLL_State".M[88, 4]) AND (NOT "ROLL_State".M[88, 5]) AND (NOT "ROLL_State".M[88, 6]));
    "ROLL_State".M[31, 2] := #r;
    // PB7, STEP 5 network 21
    #r := ("ROLL_State".M[30, 5] AND "ROLL_State".M[30, 6] AND "ROLL_State".M[30, 7] AND "ROLL_State".M[31, 0] AND "ROLL_State".M[31, 2]);
    "ROLL_State".M[31, 1] := #r;
    // PB7, STEP 5 network 22
    #r := (("ROLL_State".M[28, 4] OR "ROLL_State".M[31, 5]) AND "ROLL_IO".Input[0, 4] AND "ROLL_State".M[4, 4]);
    IF #r THEN "ROLL_State".M[31, 4] := TRUE; END_IF;
    #r := ((NOT "ROLL_IO".Input[0, 2]) OR (NOT "ROLL_IO".Input[0, 3]) OR (NOT "ROLL_State".M[29, 0]) OR (NOT "ROLL_State".M[31, 1]));
    IF #r THEN "ROLL_State".M[31, 4] := FALSE; END_IF;
    // PB7, STEP 5 network 23
    #r := "ROLL_State".M[31, 4];
    IF #r THEN "ROLL_State".M[31, 5] := TRUE; END_IF;
    #r := (((NOT "ROLL_State".M[31, 4]) AND (((NOT "ROLL_State".M[37, 2]) AND "ROLL_State".M[37, 1]) OR "ROLL_State".M[37, 0]) AND "ROLL_State".M[28, 4]) OR (NOT "ROLL_IO".Input[0, 2]));
    IF #r THEN "ROLL_State".M[31, 5] := FALSE; END_IF;
    // PB7, STEP 5 network 24
    #r := "ROLL_State".M[52, 3];
    IF #r THEN "ROLL_State".M[31, 6] := TRUE; END_IF;
    #r := ((NOT "ROLL_IO".Input[14, 0]) AND "ROLL_IO".Input[12, 1]);
    IF #r THEN "ROLL_State".M[31, 6] := FALSE; END_IF;
    // PB7, STEP 5 network 25
    #r := "ROLL_State".M[31, 5];
    "ROLL_IO".Output[16, 6] := #r;
    // PB7, STEP 5 network 26
    #r := "ROLL_State".M[40, 0];
    "ROLL_IO".Output[16, 7] := #r;
    // PB7, STEP 5 network 27
    RETURN;
END_FUNCTION

FUNCTION "ROLL_PB8" : Void
{ S7_Optimized_Access := 'TRUE' }
VERSION : 0.1
VAR_TEMP
    r : Bool;
    a1 : Word;
    a2 : Word;
    activeDataBlock : Int;
    comparisonResults : Array[0..0] of Bool;
END_VAR
BEGIN
    #r := FALSE;
    #a1 := W#16#0000;
    #a2 := W#16#0000;
    #activeDataBlock := 0;
    // PB8, STEP 5 network 1
    #r := ("ROLL_State".M[37, 7] OR "ROLL_State".M[38, 0] OR "ROLL_State".M[39, 7] OR "ROLL_State".M[40, 0] OR "ROLL_State".M[40, 1] OR "ROLL_State".M[40, 4] OR "ROLL_State".M[41, 0] OR "ROLL_State".M[41, 6] OR "ROLL_State".M[41, 7] OR "ROLL_State".M[42, 2] OR "ROLL_State".M[42, 3]);
    "ROLL_State".M[33, 0] := #r;
    // PB8, STEP 5 network 2
    #r := (((NOT "ROLL_State".M[16, 0]) AND (NOT "ROLL_State".M[16, 1]) AND (NOT "ROLL_State".M[16, 4]) AND "ROLL_State".M[37, 2]) OR "ROLL_State".M[37, 3] OR "ROLL_State".M[37, 5] OR "ROLL_State".M[37, 6] OR "ROLL_State".M[39, 4] OR "ROLL_State".M[39, 5] OR "ROLL_State".M[40, 2] OR "ROLL_State".M[40, 3] OR "ROLL_State".M[40, 6] OR "ROLL_State".M[40, 7] OR "ROLL_State".M[41, 2] OR "ROLL_State".M[42, 0] OR "ROLL_State".M[42, 4]);
    "ROLL_State".M[33, 1] := #r;
    // PB8, STEP 5 network 3
    #a2 := #a1;
    #a1 := W#16#2030;
    #r := ((NOT "ROLL_State".M[3, 1]) AND ("ROLL_State".M[33, 0] OR "ROLL_State".M[42, 6] OR "ROLL_State".M[43, 4] OR "ROLL_State".M[43, 6] OR "ROLL_State".M[43, 7] OR "ROLL_State".M[44, 2] OR "ROLL_State".M[45, 0] OR "ROLL_State".M[45, 1] OR "ROLL_State".M[45, 5] OR "ROLL_State".M[45, 7] OR "ROLL_State".M[46, 1] OR "ROLL_State".M[46, 4] OR "ROLL_State".M[46, 6] OR "ROLL_State".M[52, 1] OR "ROLL_State".M[52, 2] OR "ROLL_State".M[53, 3]) AND "ROLL_IO".Input[0, 2] AND "ROLL_State".M[29, 0]);
    "ROLL_TimerOp"(Number := 40, Operation := 0, Signal := #r, Preset := #a1);
    // PB8, STEP 5 network 4
    #a2 := #a1;
    #a1 := W#16#2030;
    #r := ((NOT "ROLL_State".M[3, 1]) AND (((NOT "ROLL_IO".Input[11, 2]) AND "ROLL_State".M[52, 0]) OR ((NOT "ROLL_State".M[15, 1]) AND "ROLL_State".M[53, 1]) OR "ROLL_State".M[33, 1] OR "ROLL_State".M[43, 0] OR "ROLL_State".M[43, 2] OR "ROLL_State".M[43, 3] OR "ROLL_State".M[44, 0] OR "ROLL_State".M[44, 7] OR "ROLL_State".M[45, 3] OR "ROLL_State".M[45, 4] OR "ROLL_State".M[46, 2] OR "ROLL_State".M[46, 3] OR "ROLL_State".M[46, 7] OR "ROLL_State".M[47, 3] OR "ROLL_State".M[52, 3] OR "ROLL_State".M[53, 2] OR "ROLL_State".M[53, 5] OR "ROLL_State".M[53, 6]) AND "ROLL_IO".Input[0, 2] AND "ROLL_State".M[29, 0]);
    "ROLL_TimerOp"(Number := 41, Operation := 0, Signal := #r, Preset := #a1);
    // PB8, STEP 5 network 5
    #r := ("ROLL_State".S5Timers[40].Q OR "ROLL_State".S5Timers[41].Q);
    IF #r THEN "ROLL_State".M[34, 1] := TRUE; END_IF;
    #r := ((NOT "ROLL_IO".Input[0, 2]) OR "ROLL_State".M[3, 1]);
    IF #r THEN "ROLL_State".M[34, 1] := FALSE; END_IF;
    // PB8, STEP 5 network 6
    RETURN;
END_FUNCTION

FUNCTION "ROLL_PB9" : Void
{ S7_Optimized_Access := 'TRUE' }
VERSION : 0.1
VAR_TEMP
    r : Bool;
    a1 : Word;
    a2 : Word;
    activeDataBlock : Int;
    comparisonResults : Array[0..0] of Bool;
END_VAR
BEGIN
    #r := FALSE;
    #a1 := W#16#0000;
    #a2 := W#16#0000;
    #activeDataBlock := 0;
    // PB9, STEP 5 network 1
    #r := ((NOT "ROLL_State".M[32, 1]) AND (NOT "ROLL_State".M[32, 2]) AND "ROLL_IO".Input[0, 2]);
    "ROLL_State".M[32, 0] := #r;
    // PB9, STEP 5 network 2
    #r := "ROLL_State".M[32, 0];
    IF #r THEN "ROLL_State".M[32, 1] := TRUE; END_IF;
    #r := ((NOT "ROLL_IO".Input[0, 2]) OR "ROLL_IO".Input[0, 1] OR "ROLL_State".M[32, 2]);
    IF #r THEN "ROLL_State".M[32, 1] := FALSE; END_IF;
    // PB9, STEP 5 network 3
    #r := ((NOT "ROLL_IO".Input[0, 2]) OR "ROLL_IO".Input[0, 1]);
    "ROLL_State".M[32, 2] := #r;
    // PB9, STEP 5 network 4
    #r := ((NOT "ROLL_State".M[12, 0]) AND (NOT "ROLL_State".M[5, 0]) AND (NOT "ROLL_State".M[5, 2]) AND (NOT "ROLL_State".M[9, 0]));
    "ROLL_State".M[35, 1] := #r;
    // PB9, STEP 5 network 5
    #r := "ROLL_IO".Input[0, 4];
    IF #r THEN "ROLL_State".M[35, 2] := TRUE; END_IF;
    #r := ((NOT "ROLL_State".M[29, 0]) OR (NOT "ROLL_State".M[31, 5]) OR (NOT "ROLL_State".M[35, 1]) OR "ROLL_State".M[16, 3]);
    IF #r THEN "ROLL_State".M[35, 2] := FALSE; END_IF;
    // PB9, STEP 5 network 6
    #r := ("ROLL_State".M[32, 0] OR "ROLL_State".M[53, 6]);
    IF #r THEN "ROLL_State".M[37, 0] := TRUE; END_IF;
    #r := ("ROLL_State".M[32, 2] OR "ROLL_State".M[37, 1] OR "ROLL_State".M[38, 0] OR "ROLL_State".M[39, 5]);
    IF #r THEN "ROLL_State".M[37, 0] := FALSE; END_IF;
    // PB9, STEP 5 network 7
    #r := ((NOT "ROLL_IO".Input[123, 5]) AND (NOT "ROLL_IO".Input[123, 6]) AND (NOT "ROLL_State".M[53, 6]) AND "ROLL_State".M[31, 5] AND "ROLL_State".M[35, 2] AND "ROLL_State".M[37, 0]);
    IF #r THEN "ROLL_State".M[37, 1] := TRUE; END_IF;
    #r := ("ROLL_State".M[32, 2] OR "ROLL_State".M[37, 2] OR "ROLL_State".M[39, 6]);
    IF #r THEN "ROLL_State".M[37, 1] := FALSE; END_IF;
    // PB9, STEP 5 network 8
    #r := ((NOT "ROLL_IO".Output[113, 3]) AND (NOT "ROLL_State".M[9, 1]) AND (("ROLL_IO".Input[0, 5] AND "ROLL_IO".Input[14, 3] AND "ROLL_State".M[0, 4]) OR ("ROLL_IO".Input[123, 4] AND "ROLL_IO".Input[124, 4] AND "ROLL_State".M[0, 3])) AND "ROLL_State".M[35, 2] AND "ROLL_State".M[37, 1]);
    IF #r THEN "ROLL_State".M[37, 2] := TRUE; END_IF;
    #r := ("ROLL_State".M[32, 2] OR "ROLL_State".M[37, 3]);
    IF #r THEN "ROLL_State".M[37, 2] := FALSE; END_IF;
    // PB9, STEP 5 network 9
    #r := ((NOT "ROLL_State".M[16, 0]) AND (NOT "ROLL_State".M[16, 1]) AND (NOT "ROLL_State".M[16, 4]) AND (NOT "ROLL_State".M[191, 5]) AND "ROLL_IO".Input[14, 0] AND "ROLL_State".M[190, 1] AND "ROLL_State".M[191, 4] AND "ROLL_State".M[35, 2] AND "ROLL_State".M[37, 2]);
    IF #r THEN "ROLL_State".M[37, 3] := TRUE; END_IF;
    #r := ("ROLL_State".M[32, 2] OR "ROLL_State".M[37, 5] OR "ROLL_State".M[40, 0]);
    IF #r THEN "ROLL_State".M[37, 3] := FALSE; END_IF;
    // PB9, STEP 5 network 10
    #r := ((NOT "ROLL_IO".Input[123, 5]) AND (NOT "ROLL_IO".Input[123, 6]) AND "ROLL_IO".Input[124, 1] AND "ROLL_IO".Input[124, 4] AND "ROLL_State".M[0, 3] AND "ROLL_State".M[35, 2] AND "ROLL_State".M[37, 3]);
    IF #r THEN "ROLL_State".M[37, 5] := TRUE; END_IF;
    #r := ("ROLL_State".M[32, 2] OR "ROLL_State".M[37, 6]);
    IF #r THEN "ROLL_State".M[37, 5] := FALSE; END_IF;
    // PB9, STEP 5 network 11
    #r := ((NOT "ROLL_IO".Output[113, 2]) AND "ROLL_IO".Output[113, 3] AND "ROLL_State".M[35, 2] AND "ROLL_State".M[37, 5] AND "ROLL_State".S5Timers[18].Q);
    IF #r THEN "ROLL_State".M[37, 6] := TRUE; END_IF;
    #r := ("ROLL_State".M[32, 2] OR "ROLL_State".M[37, 7]);
    IF #r THEN "ROLL_State".M[37, 6] := FALSE; END_IF;
    // PB9, STEP 5 network 12
    #r := ((NOT "ROLL_State".M[37, 5]) AND "ROLL_State".M[35, 2] AND "ROLL_State".M[37, 6]);
    IF #r THEN "ROLL_State".M[37, 7] := TRUE; END_IF;
    #r := ("ROLL_State".M[32, 2] OR "ROLL_State".M[38, 0]);
    IF #r THEN "ROLL_State".M[37, 7] := FALSE; END_IF;
    // PB9, STEP 5 network 13
    #r := ((NOT "ROLL_State".M[70, 2]) AND (((NOT "ROLL_IO".Output[113, 2]) AND "ROLL_IO".Output[113, 3] AND "ROLL_IO".Input[124, 4] AND "ROLL_State".M[28, 4] AND "ROLL_State".M[37, 0]) OR ("ROLL_State".M[37, 7] AND "ROLL_State".S5Timers[20].Q)) AND "ROLL_IO".Input[123, 5] AND "ROLL_State".M[35, 2]);
    IF #r THEN "ROLL_State".M[38, 0] := TRUE; END_IF;
    #r := ("ROLL_State".M[32, 2] OR "ROLL_State".M[39, 4]);
    IF #r THEN "ROLL_State".M[38, 0] := FALSE; END_IF;
    // PB9, STEP 5 network 14
    #r := ((NOT "ROLL_IO".Input[124, 5]) AND "ROLL_IO".Input[124, 4] AND "ROLL_State".M[35, 2] AND "ROLL_State".M[38, 0]);
    IF #r THEN "ROLL_State".M[39, 4] := TRUE; END_IF;
    #r := ("ROLL_State".M[32, 2] OR "ROLL_State".M[39, 5]);
    IF #r THEN "ROLL_State".M[39, 4] := FALSE; END_IF;
    // PB9, STEP 5 network 15
    #r := ((NOT "ROLL_IO".Input[124, 4]) AND (("ROLL_State".M[28, 4] AND "ROLL_State".M[37, 0]) OR "ROLL_State".M[39, 4]) AND "ROLL_IO".Input[124, 5] AND "ROLL_State".M[35, 2]);
    IF #r THEN "ROLL_State".M[39, 5] := TRUE; END_IF;
    #r := ("ROLL_State".M[32, 2] OR "ROLL_State".M[39, 6]);
    IF #r THEN "ROLL_State".M[39, 5] := FALSE; END_IF;
    // PB9, STEP 5 network 16
    #r := ((NOT "ROLL_IO".Input[124, 2]) AND "ROLL_IO".Input[11, 0] AND "ROLL_IO".Input[11, 6] AND "ROLL_IO".Input[12, 1] AND "ROLL_IO".Input[12, 7] AND "ROLL_IO".Input[124, 1] AND "ROLL_State".M[35, 2] AND "ROLL_State".M[39, 5]);
    IF #r THEN "ROLL_State".M[39, 6] := TRUE; END_IF;
    #r := ("ROLL_State".M[32, 2] OR "ROLL_State".M[39, 7]);
    IF #r THEN "ROLL_State".M[39, 6] := FALSE; END_IF;
    // PB9, STEP 5 network 17
    #r := ((NOT "ROLL_IO".Input[124, 1]) AND "ROLL_IO".Input[124, 2] AND "ROLL_State".M[35, 2] AND "ROLL_State".M[39, 6]);
    IF #r THEN "ROLL_State".M[39, 7] := TRUE; END_IF;
    #r := ("ROLL_State".M[32, 2] OR "ROLL_State".M[40, 0]);
    IF #r THEN "ROLL_State".M[39, 7] := FALSE; END_IF;
    // PB9, STEP 5 network 18
    #r := ((NOT "ROLL_IO".Input[12, 5]) AND ("ROLL_State".M[37, 3] OR "ROLL_State".M[39, 7]) AND "ROLL_IO".Input[11, 0] AND "ROLL_IO".Input[11, 6] AND "ROLL_IO".Input[12, 1] AND "ROLL_IO".Input[12, 7] AND "ROLL_State".M[35, 2]);
    IF #r THEN "ROLL_State".M[40, 0] := TRUE; END_IF;
    #r := ("ROLL_State".M[32, 2] OR "ROLL_State".M[40, 1]);
    IF #r THEN "ROLL_State".M[40, 0] := FALSE; END_IF;
    // PB9, STEP 5 network 19
    #r := ("ROLL_IO".Input[12, 5] AND "ROLL_IO".Input[12, 7] AND "ROLL_State".M[35, 2] AND "ROLL_State".M[40, 0]);
    IF #r THEN "ROLL_State".M[40, 1] := TRUE; END_IF;
    #r := ("ROLL_State".M[32, 2] OR "ROLL_State".M[40, 2] OR "ROLL_State".M[41, 6] OR "ROLL_State".M[43, 2] OR "ROLL_State".M[44, 7] OR "ROLL_State".M[46, 2] OR "ROLL_State".M[47, 6] OR "ROLL_State".M[49, 2] OR "ROLL_State".M[50, 6]);
    IF #r THEN "ROLL_State".M[40, 1] := FALSE; END_IF;
    // PB9, STEP 5 network 20
    #r := ((NOT "ROLL_IO".Input[11, 1]) AND "ROLL_IO".Input[11, 0] AND "ROLL_State".M[110, 0] AND "ROLL_State".M[35, 2] AND "ROLL_State".M[40, 1] AND "ROLL_State".M[63, 1]);
    IF #r THEN "ROLL_State".M[40, 2] := TRUE; END_IF;
    #r := ("ROLL_State".M[32, 2] OR "ROLL_State".M[40, 3]);
    IF #r THEN "ROLL_State".M[40, 2] := FALSE; END_IF;
    // PB9, STEP 5 network 21
    #r := ("ROLL_IO".Input[11, 1] AND "ROLL_IO".Input[11, 6] AND "ROLL_State".M[35, 2] AND "ROLL_State".M[40, 2]);
    IF #r THEN "ROLL_State".M[40, 3] := TRUE; END_IF;
    #r := ("ROLL_State".M[32, 2] OR "ROLL_State".M[40, 4]);
    IF #r THEN "ROLL_State".M[40, 3] := FALSE; END_IF;
    // PB9, STEP 5 network 22
    #r := ((NOT "ROLL_IO".Input[12, 1]) AND "ROLL_IO".Input[12, 5] AND "ROLL_State".M[35, 2] AND "ROLL_State".M[40, 3]);
    IF #r THEN "ROLL_State".M[40, 4] := TRUE; END_IF;
    #r := ("ROLL_State".M[32, 2] OR "ROLL_State".M[40, 5]);
    IF #r THEN "ROLL_State".M[40, 4] := FALSE; END_IF;
    // PB9, STEP 5 network 23
    #r := ("ROLL_IO".Input[12, 1] AND "ROLL_IO".Input[12, 7] AND "ROLL_State".M[35, 2] AND "ROLL_State".M[40, 4]);
    IF #r THEN "ROLL_State".M[40, 5] := TRUE; END_IF;
    #r := ("ROLL_State".M[32, 2] OR "ROLL_State".M[40, 6]);
    IF #r THEN "ROLL_State".M[40, 5] := FALSE; END_IF;
    // PB9, STEP 5 network 24
    #r := ("ROLL_State".M[35, 2] AND "ROLL_State".M[40, 5] AND "ROLL_State".S5Timers[1].Q);
    IF #r THEN "ROLL_State".M[40, 6] := TRUE; END_IF;
    #r := ("ROLL_State".M[32, 2] OR "ROLL_State".M[40, 7]);
    IF #r THEN "ROLL_State".M[40, 6] := FALSE; END_IF;
    // PB9, STEP 5 network 25
    #r := ("ROLL_State".M[35, 2] AND "ROLL_State".M[40, 6]);
    IF #r THEN "ROLL_State".M[40, 7] := TRUE; END_IF;
    #r := ("ROLL_State".M[32, 2] OR "ROLL_State".M[41, 0]);
    IF #r THEN "ROLL_State".M[40, 7] := FALSE; END_IF;
    // PB9, STEP 5 network 26
    #r := ((NOT "ROLL_IO".Input[12, 5]) AND (("ROLL_IO".Input[13, 3] AND "ROLL_State".M[63, 1]) OR (NOT "ROLL_State".M[111, 5])) AND "ROLL_State".M[35, 2] AND "ROLL_State".M[40, 7]);
    IF #r THEN "ROLL_State".M[41, 0] := TRUE; END_IF;
    #r := ("ROLL_State".M[32, 2] OR "ROLL_State".M[41, 1]);
    IF #r THEN "ROLL_State".M[41, 0] := FALSE; END_IF;
    // PB9, STEP 5 network 27
    #r := ("ROLL_IO".Input[12, 5] AND "ROLL_IO".Input[12, 7] AND "ROLL_State".M[35, 2] AND "ROLL_State".M[41, 0]);
    IF #r THEN "ROLL_State".M[41, 1] := TRUE; END_IF;
    #r := ("ROLL_State".M[32, 2] OR "ROLL_State".M[41, 2]);
    IF #r THEN "ROLL_State".M[41, 1] := FALSE; END_IF;
    // PB9, STEP 5 network 28
    #r := ("ROLL_State".M[35, 2] AND "ROLL_State".M[41, 1] AND "ROLL_State".S5Timers[2].Q);
    IF #r THEN "ROLL_State".M[41, 2] := TRUE; END_IF;
    #r := ("ROLL_State".M[32, 2] OR "ROLL_State".M[41, 3] OR "ROLL_State".M[41, 6] OR "ROLL_State".M[43, 2] OR "ROLL_State".M[44, 7] OR "ROLL_State".M[46, 2] OR "ROLL_State".M[47, 6] OR "ROLL_State".M[49, 2]);
    IF #r THEN "ROLL_State".M[41, 2] := FALSE; END_IF;
    // PB9, STEP 5 network 29
    #r := ((NOT "ROLL_State".M[110, 1]) AND (NOT "ROLL_State".M[110, 2]) AND "ROLL_State".M[35, 2] AND "ROLL_State".M[41, 2]);
    IF #r THEN "ROLL_State".M[41, 3] := TRUE; END_IF;
    #r := ("ROLL_State".M[32, 2] OR "ROLL_State".M[41, 4]);
    IF #r THEN "ROLL_State".M[41, 3] := FALSE; END_IF;
    // PB9, STEP 5 network 30
    #r := ("ROLL_IO".Input[13, 3] AND "ROLL_State".M[35, 2] AND "ROLL_State".M[41, 3] AND "ROLL_State".M[63, 1]);
    IF #r THEN "ROLL_State".M[41, 4] := TRUE; END_IF;
    #r := ("ROLL_State".M[32, 2] OR "ROLL_State".M[44, 7] OR "ROLL_State".M[50, 6] OR "ROLL_State".M[52, 0]);
    IF #r THEN "ROLL_State".M[41, 4] := FALSE; END_IF;
    // PB9, STEP 5 network 31
    #r := ((NOT "ROLL_IO".Input[11, 2]) AND (((NOT "ROLL_State".M[110, 0]) AND "ROLL_State".M[40, 1]) OR "ROLL_State".M[41, 2]) AND "ROLL_IO".Input[12, 5] AND "ROLL_IO".Input[12, 7] AND "ROLL_State".M[110, 1] AND "ROLL_State".M[35, 2]);
    IF #r THEN "ROLL_State".M[41, 6] := TRUE; END_IF;
    #r := ("ROLL_State".M[32, 2] OR "ROLL_State".M[41, 7]);
    IF #r THEN "ROLL_State".M[41, 6] := FALSE; END_IF;
    // PB9, STEP 5 network 32
    #r := ("ROLL_IO".Input[11, 2] AND "ROLL_IO".Input[11, 6] AND "ROLL_State".M[35, 2] AND "ROLL_State".M[41, 6]);
    IF #r THEN "ROLL_State".M[41, 7] := TRUE; END_IF;
    #r := ("ROLL_State".M[32, 2] OR "ROLL_State".M[42, 0]);
    IF #r THEN "ROLL_State".M[41, 7] := FALSE; END_IF;
    // PB9, STEP 5 network 33
    #r := ((NOT "ROLL_IO".Input[12, 1]) AND "ROLL_IO".Input[12, 5] AND "ROLL_State".M[35, 2] AND "ROLL_State".M[41, 7]);
    IF #r THEN "ROLL_State".M[42, 0] := TRUE; END_IF;
    #r := ("ROLL_State".M[32, 2] OR "ROLL_State".M[42, 1]);
    IF #r THEN "ROLL_State".M[42, 0] := FALSE; END_IF;
    // PB9, STEP 5 network 34
    #r := ("ROLL_IO".Input[12, 1] AND "ROLL_IO".Input[12, 7] AND "ROLL_State".M[35, 2] AND "ROLL_State".M[42, 0]);
    IF #r THEN "ROLL_State".M[42, 1] := TRUE; END_IF;
    #r := ("ROLL_State".M[32, 2] OR "ROLL_State".M[42, 2]);
    IF #r THEN "ROLL_State".M[42, 1] := FALSE; END_IF;
    // PB9, STEP 5 network 35
    #r := ("ROLL_State".M[35, 2] AND "ROLL_State".M[42, 1] AND "ROLL_State".S5Timers[1].Q);
    IF #r THEN "ROLL_State".M[42, 2] := TRUE; END_IF;
    #r := ("ROLL_State".M[32, 2] OR "ROLL_State".M[42, 3]);
    IF #r THEN "ROLL_State".M[42, 2] := FALSE; END_IF;
    // PB9, STEP 5 network 36
    #r := ("ROLL_State".M[35, 2] AND "ROLL_State".M[42, 2]);
    IF #r THEN "ROLL_State".M[42, 3] := TRUE; END_IF;
    #r := ("ROLL_State".M[32, 2] OR "ROLL_State".M[42, 4]);
    IF #r THEN "ROLL_State".M[42, 3] := FALSE; END_IF;
    // PB9, STEP 5 network 37
    #r := ((NOT "ROLL_IO".Input[12, 5]) AND (("ROLL_IO".Input[13, 3] AND "ROLL_State".M[63, 1]) OR (NOT "ROLL_State".M[111, 5])) AND "ROLL_State".M[35, 2] AND "ROLL_State".M[42, 3]);
    IF #r THEN "ROLL_State".M[42, 4] := TRUE; END_IF;
    #r := ("ROLL_State".M[32, 2] OR "ROLL_State".M[42, 5]);
    IF #r THEN "ROLL_State".M[42, 4] := FALSE; END_IF;
    // PB9, STEP 5 network 38
    #r := ("ROLL_IO".Input[12, 5] AND "ROLL_IO".Input[12, 7] AND "ROLL_State".M[35, 2] AND "ROLL_State".M[42, 4]);
    IF #r THEN "ROLL_State".M[42, 5] := TRUE; END_IF;
    #r := ("ROLL_State".M[32, 2] OR "ROLL_State".M[42, 6]);
    IF #r THEN "ROLL_State".M[42, 5] := FALSE; END_IF;
    // PB9, STEP 5 network 39
    #r := ("ROLL_State".M[35, 2] AND "ROLL_State".M[42, 5] AND "ROLL_State".S5Timers[2].Q);
    IF #r THEN "ROLL_State".M[42, 6] := TRUE; END_IF;
    #r := ("ROLL_State".M[32, 2] OR "ROLL_State".M[42, 7] OR "ROLL_State".M[43, 2] OR "ROLL_State".M[44, 7] OR "ROLL_State".M[46, 2] OR "ROLL_State".M[47, 6] OR "ROLL_State".M[49, 2]);
    IF #r THEN "ROLL_State".M[42, 6] := FALSE; END_IF;
    // PB9, STEP 5 network 40
    #r := ((NOT "ROLL_State".M[110, 2]) AND "ROLL_State".M[35, 2] AND "ROLL_State".M[42, 6]);
    IF #r THEN "ROLL_State".M[42, 7] := TRUE; END_IF;
    #r := ("ROLL_State".M[32, 2] OR "ROLL_State".M[43, 0]);
    IF #r THEN "ROLL_State".M[42, 7] := FALSE; END_IF;
    // PB9, STEP 5 network 41
    #r := ("ROLL_IO".Input[13, 3] AND "ROLL_State".M[35, 2] AND "ROLL_State".M[42, 7] AND "ROLL_State".M[63, 1]);
    IF #r THEN "ROLL_State".M[43, 0] := TRUE; END_IF;
    #r := ("ROLL_State".M[32, 2] OR "ROLL_State".M[44, 7] OR "ROLL_State".M[50, 6] OR "ROLL_State".M[52, 0]);
    IF #r THEN "ROLL_State".M[43, 0] := FALSE; END_IF;
    // PB9, STEP 5 network 42
    #r := ((NOT "ROLL_IO".Input[11, 3]) AND (((NOT "ROLL_State".M[110, 0]) AND (NOT "ROLL_State".M[110, 1]) AND "ROLL_State".M[40, 1]) OR ((NOT "ROLL_State".M[110, 1]) AND "ROLL_State".M[41, 2]) OR "ROLL_State".M[42, 6]) AND "ROLL_IO".Input[12, 5] AND "ROLL_IO".Input[12, 7] AND "ROLL_State".M[110, 2] AND "ROLL_State".M[35, 2]);
    IF #r THEN "ROLL_State".M[43, 2] := TRUE; END_IF;
    #r := ("ROLL_State".M[32, 2] OR "ROLL_State".M[43, 3]);
    IF #r THEN "ROLL_State".M[43, 2] := FALSE; END_IF;
    // PB9, STEP 5 network 43
    #r := ("ROLL_IO".Input[11, 3] AND "ROLL_IO".Input[11, 6] AND "ROLL_State".M[35, 2] AND "ROLL_State".M[43, 2]);
    IF #r THEN "ROLL_State".M[43, 3] := TRUE; END_IF;
    #r := ("ROLL_State".M[32, 2] OR "ROLL_State".M[43, 4]);
    IF #r THEN "ROLL_State".M[43, 3] := FALSE; END_IF;
    // PB9, STEP 5 network 44
    #r := ((NOT "ROLL_IO".Input[12, 1]) AND "ROLL_IO".Input[12, 5] AND "ROLL_State".M[35, 2] AND "ROLL_State".M[43, 3]);
    IF #r THEN "ROLL_State".M[43, 4] := TRUE; END_IF;
    #r := ("ROLL_State".M[32, 2] OR "ROLL_State".M[43, 5]);
    IF #r THEN "ROLL_State".M[43, 4] := FALSE; END_IF;
    // PB9, STEP 5 network 45
    #r := ("ROLL_IO".Input[12, 1] AND "ROLL_IO".Input[12, 7] AND "ROLL_State".M[35, 2] AND "ROLL_State".M[43, 4]);
    IF #r THEN "ROLL_State".M[43, 5] := TRUE; END_IF;
    #r := ("ROLL_State".M[32, 2] OR "ROLL_State".M[43, 6]);
    IF #r THEN "ROLL_State".M[43, 5] := FALSE; END_IF;
    // PB9, STEP 5 network 46
    #r := ("ROLL_State".M[35, 2] AND "ROLL_State".M[43, 5] AND "ROLL_State".S5Timers[1].Q);
    IF #r THEN "ROLL_State".M[43, 6] := TRUE; END_IF;
    #r := ("ROLL_State".M[32, 2] OR "ROLL_State".M[43, 7]);
    IF #r THEN "ROLL_State".M[43, 6] := FALSE; END_IF;
    // PB9, STEP 5 network 47
    #r := ("ROLL_State".M[35, 2] AND "ROLL_State".M[43, 6]);
    IF #r THEN "ROLL_State".M[43, 7] := TRUE; END_IF;
    #r := ("ROLL_State".M[32, 2] OR "ROLL_State".M[44, 0]);
    IF #r THEN "ROLL_State".M[43, 7] := FALSE; END_IF;
    // PB9, STEP 5 network 48
    #r := ((NOT "ROLL_IO".Input[12, 5]) AND (("ROLL_IO".Input[13, 3] AND "ROLL_State".M[63, 1]) OR (NOT "ROLL_State".M[111, 5])) AND "ROLL_State".M[35, 2] AND "ROLL_State".M[43, 7]);
    IF #r THEN "ROLL_State".M[44, 0] := TRUE; END_IF;
    #r := ("ROLL_State".M[32, 2] OR "ROLL_State".M[44, 1]);
    IF #r THEN "ROLL_State".M[44, 0] := FALSE; END_IF;
    // PB9, STEP 5 network 49
    #r := ("ROLL_IO".Input[12, 5] AND "ROLL_IO".Input[12, 7] AND "ROLL_State".M[35, 2] AND "ROLL_State".M[44, 0]);
    IF #r THEN "ROLL_State".M[44, 1] := TRUE; END_IF;
    #r := ("ROLL_State".M[32, 2] OR "ROLL_State".M[44, 2]);
    IF #r THEN "ROLL_State".M[44, 1] := FALSE; END_IF;
    // PB9, STEP 5 network 50
    #r := ("ROLL_State".M[35, 2] AND "ROLL_State".M[44, 1] AND "ROLL_State".S5Timers[2].Q);
    IF #r THEN "ROLL_State".M[44, 2] := TRUE; END_IF;
    #r := ("ROLL_State".M[32, 2] OR "ROLL_State".M[44, 3] OR "ROLL_State".M[44, 7] OR "ROLL_State".M[46, 2] OR "ROLL_State".M[47, 6] OR "ROLL_State".M[49, 2]);
    IF #r THEN "ROLL_State".M[44, 2] := FALSE; END_IF;
    // PB9, STEP 5 network 51
    #r := ("ROLL_State".M[35, 2] AND "ROLL_State".M[44, 2]);
    IF #r THEN "ROLL_State".M[44, 3] := TRUE; END_IF;
    #r := ("ROLL_State".M[32, 2] OR "ROLL_State".M[44, 4]);
    IF #r THEN "ROLL_State".M[44, 3] := FALSE; END_IF;
    // PB9, STEP 5 network 52
    #r := ("ROLL_IO".Input[13, 3] AND "ROLL_State".M[35, 2] AND "ROLL_State".M[44, 3] AND "ROLL_State".M[63, 1]);
    IF #r THEN "ROLL_State".M[44, 4] := TRUE; END_IF;
    #r := ("ROLL_State".M[32, 2] OR "ROLL_State".M[44, 7] OR "ROLL_State".M[50, 6] OR "ROLL_State".M[52, 0]);
    IF #r THEN "ROLL_State".M[44, 4] := FALSE; END_IF;
    // PB9, STEP 5 network 53
    #r := (((NOT "ROLL_State".M[110, 0]) AND (NOT "ROLL_State".M[110, 1]) AND (NOT "ROLL_State".M[110, 2]) AND "ROLL_State".M[40, 1]) OR ((NOT "ROLL_State".M[110, 1]) AND (NOT "ROLL_State".M[110, 2]) AND "ROLL_State".M[41, 4]) OR ((NOT "ROLL_State".M[110, 2]) AND "ROLL_State".M[43, 0]) OR "ROLL_State".M[44, 4]);
    "ROLL_State".M[240, 0] := #r;
    // PB9, STEP 5 network 54
    #r := ((NOT "ROLL_IO".Input[11, 4]) AND "ROLL_IO".Input[12, 5] AND "ROLL_IO".Input[12, 7] AND "ROLL_State".M[110, 3] AND "ROLL_State".M[240, 0] AND "ROLL_State".M[35, 2] AND "ROLL_State".M[63, 1]);
    IF #r THEN "ROLL_State".M[44, 7] := TRUE; END_IF;
    #r := ("ROLL_State".M[32, 2] OR "ROLL_State".M[45, 0]);
    IF #r THEN "ROLL_State".M[44, 7] := FALSE; END_IF;
    // PB9, STEP 5 network 55
    #r := ("ROLL_IO".Input[11, 4] AND "ROLL_IO".Input[11, 6] AND "ROLL_State".M[35, 2] AND "ROLL_State".M[44, 7]);
    IF #r THEN "ROLL_State".M[45, 0] := TRUE; END_IF;
    #r := ("ROLL_State".M[32, 2] OR "ROLL_State".M[45, 1]);
    IF #r THEN "ROLL_State".M[45, 0] := FALSE; END_IF;
    // PB9, STEP 5 network 56
    #r := ((NOT "ROLL_IO".Input[12, 1]) AND "ROLL_IO".Input[12, 5] AND "ROLL_State".M[35, 2] AND "ROLL_State".M[45, 0]);
    IF #r THEN "ROLL_State".M[45, 1] := TRUE; END_IF;
    #r := ("ROLL_State".M[32, 2] OR "ROLL_State".M[45, 2]);
    IF #r THEN "ROLL_State".M[45, 1] := FALSE; END_IF;
    // PB9, STEP 5 network 57
    #r := ("ROLL_IO".Input[12, 1] AND "ROLL_IO".Input[12, 7] AND "ROLL_State".M[35, 2] AND "ROLL_State".M[45, 1]);
    IF #r THEN "ROLL_State".M[45, 2] := TRUE; END_IF;
    #r := ("ROLL_State".M[32, 2] OR "ROLL_State".M[45, 3]);
    IF #r THEN "ROLL_State".M[45, 2] := FALSE; END_IF;
    // PB9, STEP 5 network 58
    #r := ("ROLL_State".M[35, 2] AND "ROLL_State".M[45, 2] AND "ROLL_State".S5Timers[1].Q);
    IF #r THEN "ROLL_State".M[45, 3] := TRUE; END_IF;
    #r := ("ROLL_State".M[32, 2] OR "ROLL_State".M[45, 4]);
    IF #r THEN "ROLL_State".M[45, 3] := FALSE; END_IF;
    // PB9, STEP 5 network 59
    #r := ("ROLL_State".M[35, 2] AND "ROLL_State".M[45, 3]);
    IF #r THEN "ROLL_State".M[45, 4] := TRUE; END_IF;
    #r := ("ROLL_State".M[32, 2] OR "ROLL_State".M[45, 5]);
    IF #r THEN "ROLL_State".M[45, 4] := FALSE; END_IF;
    // PB9, STEP 5 network 60
    #r := ((NOT "ROLL_IO".Input[12, 5]) AND "ROLL_State".M[35, 2] AND "ROLL_State".M[45, 4]);
    IF #r THEN "ROLL_State".M[45, 5] := TRUE; END_IF;
    #r := ("ROLL_State".M[32, 2] OR "ROLL_State".M[45, 6]);
    IF #r THEN "ROLL_State".M[45, 5] := FALSE; END_IF;
    // PB9, STEP 5 network 61
    #r := ("ROLL_IO".Input[12, 5] AND "ROLL_IO".Input[12, 7] AND "ROLL_State".M[35, 2] AND "ROLL_State".M[45, 5]);
    IF #r THEN "ROLL_State".M[45, 6] := TRUE; END_IF;
    #r := ("ROLL_State".M[32, 2] OR "ROLL_State".M[45, 7]);
    IF #r THEN "ROLL_State".M[45, 6] := FALSE; END_IF;
    // PB9, STEP 5 network 62
    #r := (("ROLL_State".M[0, 4] OR "ROLL_State".S5Timers[2].Q) AND "ROLL_State".M[35, 2] AND "ROLL_State".M[45, 6]);
    IF #r THEN "ROLL_State".M[45, 7] := TRUE; END_IF;
    #r := ("ROLL_State".M[32, 2] OR "ROLL_State".M[46, 0] OR "ROLL_State".M[46, 2] OR "ROLL_State".M[47, 6] OR "ROLL_State".M[49, 2]);
    IF #r THEN "ROLL_State".M[45, 7] := FALSE; END_IF;
    // PB9, STEP 5 network 63
    #r := ("ROLL_State".M[35, 2] AND "ROLL_State".M[45, 7]);
    IF #r THEN "ROLL_State".M[46, 0] := TRUE; END_IF;
    #r := ("ROLL_State".M[32, 2] OR "ROLL_State".M[46, 1]);
    IF #r THEN "ROLL_State".M[46, 0] := FALSE; END_IF;
    // PB9, STEP 5 network 64
    #r := ("ROLL_IO".Input[13, 3] AND "ROLL_State".M[35, 2] AND "ROLL_State".M[46, 0] AND "ROLL_State".M[63, 1]);
    IF #r THEN "ROLL_State".M[46, 1] := TRUE; END_IF;
    #r := ("ROLL_State".M[32, 2] OR "ROLL_State".M[50, 6] OR "ROLL_State".M[52, 0]);
    IF #r THEN "ROLL_State".M[46, 1] := FALSE; END_IF;
    // PB9, STEP 5 network 65
    RETURN;
END_FUNCTION

FUNCTION "ROLL_PB10" : Void
{ S7_Optimized_Access := 'TRUE' }
VERSION : 0.1
VAR_TEMP
    r : Bool;
    a1 : Word;
    a2 : Word;
    activeDataBlock : Int;
    comparisonResults : Array[0..0] of Bool;
END_VAR
BEGIN
    #r := FALSE;
    #a1 := W#16#0000;
    #a2 := W#16#0000;
    #activeDataBlock := 0;
    // PB10, STEP 5 network 1
    #r := (((NOT "ROLL_State".M[110, 0]) AND (NOT "ROLL_State".M[110, 1]) AND (NOT "ROLL_State".M[110, 2]) AND (NOT "ROLL_State".M[110, 3]) AND "ROLL_State".M[40, 1]) OR ((NOT "ROLL_State".M[110, 1]) AND (NOT "ROLL_State".M[110, 2]) AND (NOT "ROLL_State".M[110, 3]) AND "ROLL_State".M[41, 2]) OR ((NOT "ROLL_State".M[110, 2]) AND (NOT "ROLL_State".M[110, 3]) AND "ROLL_State".M[42, 6]) OR ((NOT "ROLL_State".M[110, 3]) AND "ROLL_State".M[44, 2]) OR "ROLL_State".M[45, 7]);
    "ROLL_State".M[240, 0] := #r;
    // PB10, STEP 5 network 2
    #r := ((NOT "ROLL_IO".Input[119, 6]) AND "ROLL_IO".Input[12, 5] AND "ROLL_IO".Input[12, 7] AND "ROLL_State".M[110, 4] AND "ROLL_State".M[240, 0] AND "ROLL_State".M[35, 2]);
    IF #r THEN "ROLL_State".M[46, 2] := TRUE; END_IF;
    #r := ("ROLL_State".M[32, 2] OR "ROLL_State".M[46, 3]);
    IF #r THEN "ROLL_State".M[46, 2] := FALSE; END_IF;
    // PB10, STEP 5 network 3
    #r := ("ROLL_IO".Input[11, 6] AND "ROLL_IO".Input[119, 6] AND "ROLL_State".M[35, 2] AND "ROLL_State".M[46, 2]);
    IF #r THEN "ROLL_State".M[46, 3] := TRUE; END_IF;
    #r := ("ROLL_State".M[32, 2] OR "ROLL_State".M[46, 4]);
    IF #r THEN "ROLL_State".M[46, 3] := FALSE; END_IF;
    // PB10, STEP 5 network 4
    #r := ((NOT "ROLL_IO".Input[12, 1]) AND "ROLL_IO".Input[12, 5] AND "ROLL_State".M[35, 2] AND "ROLL_State".M[46, 3]);
    IF #r THEN "ROLL_State".M[46, 4] := TRUE; END_IF;
    #r := ("ROLL_State".M[32, 2] OR "ROLL_State".M[46, 5]);
    IF #r THEN "ROLL_State".M[46, 4] := FALSE; END_IF;
    // PB10, STEP 5 network 5
    #r := ("ROLL_IO".Input[12, 1] AND "ROLL_IO".Input[12, 7] AND "ROLL_State".M[35, 2] AND "ROLL_State".M[46, 4]);
    IF #r THEN "ROLL_State".M[46, 5] := TRUE; END_IF;
    #r := ("ROLL_State".M[32, 2] OR "ROLL_State".M[46, 6]);
    IF #r THEN "ROLL_State".M[46, 5] := FALSE; END_IF;
    // PB10, STEP 5 network 6
    #r := ("ROLL_State".M[35, 2] AND "ROLL_State".M[46, 5] AND "ROLL_State".S5Timers[1].Q);
    IF #r THEN "ROLL_State".M[46, 6] := TRUE; END_IF;
    #r := ("ROLL_State".M[32, 2] OR "ROLL_State".M[46, 7]);
    IF #r THEN "ROLL_State".M[46, 6] := FALSE; END_IF;
    // PB10, STEP 5 network 7
    #r := ("ROLL_State".M[35, 2] AND "ROLL_State".M[46, 6]);
    IF #r THEN "ROLL_State".M[46, 7] := TRUE; END_IF;
    #r := ("ROLL_State".M[32, 2] OR "ROLL_State".M[47, 0]);
    IF #r THEN "ROLL_State".M[46, 7] := FALSE; END_IF;
    // PB10, STEP 5 network 8
    #r := ((NOT "ROLL_IO".Input[12, 5]) AND "ROLL_State".M[35, 2] AND "ROLL_State".M[46, 7]);
    IF #r THEN "ROLL_State".M[47, 0] := TRUE; END_IF;
    #r := ("ROLL_State".M[32, 2] OR "ROLL_State".M[47, 1]);
    IF #r THEN "ROLL_State".M[47, 0] := FALSE; END_IF;
    // PB10, STEP 5 network 9
    #r := ("ROLL_IO".Input[12, 5] AND "ROLL_IO".Input[12, 7] AND "ROLL_State".M[35, 2] AND "ROLL_State".M[47, 0]);
    IF #r THEN "ROLL_State".M[47, 1] := TRUE; END_IF;
    #r := ("ROLL_State".M[32, 2] OR "ROLL_State".M[47, 2]);
    IF #r THEN "ROLL_State".M[47, 1] := FALSE; END_IF;
    // PB10, STEP 5 network 10
    #r := ("ROLL_State".M[35, 2] AND "ROLL_State".M[47, 1] AND "ROLL_State".S5Timers[2].Q);
    IF #r THEN "ROLL_State".M[47, 2] := TRUE; END_IF;
    #r := ("ROLL_State".M[32, 2] OR "ROLL_State".M[47, 3] OR "ROLL_State".M[47, 6]);
    IF #r THEN "ROLL_State".M[47, 2] := FALSE; END_IF;
    // PB10, STEP 5 network 11
    #r := ((NOT "ROLL_State".M[110, 5]) AND (NOT "ROLL_State".M[110, 6]) AND "ROLL_State".M[35, 2] AND "ROLL_State".M[47, 2]);
    IF #r THEN "ROLL_State".M[47, 3] := TRUE; END_IF;
    #r := ("ROLL_State".M[32, 2] OR "ROLL_State".M[47, 4]);
    IF #r THEN "ROLL_State".M[47, 3] := FALSE; END_IF;
    // PB10, STEP 5 network 12
    #r := ("ROLL_IO".Input[13, 3] AND "ROLL_State".M[35, 2] AND "ROLL_State".M[47, 3] AND "ROLL_State".M[63, 1]);
    IF #r THEN "ROLL_State".M[47, 4] := TRUE; END_IF;
    #r := ("ROLL_State".M[32, 2] OR "ROLL_State".M[50, 6] OR "ROLL_State".M[52, 0]);
    IF #r THEN "ROLL_State".M[47, 4] := FALSE; END_IF;
    // PB10, STEP 5 network 13
    #r := (((NOT "ROLL_State".M[110, 0]) AND (NOT "ROLL_State".M[110, 1]) AND (NOT "ROLL_State".M[110, 2]) AND (NOT "ROLL_State".M[110, 3]) AND (NOT "ROLL_State".M[110, 4]) AND "ROLL_State".M[40, 1]) OR ((NOT "ROLL_State".M[110, 1]) AND (NOT "ROLL_State".M[110, 2]) AND (NOT "ROLL_State".M[110, 3]) AND (NOT "ROLL_State".M[110, 4]) AND "ROLL_State".M[41, 2]) OR ((NOT "ROLL_State".M[110, 2]) AND (NOT "ROLL_State".M[110, 3]) AND (NOT "ROLL_State".M[110, 4]) AND "ROLL_State".M[42, 6]) OR ((NOT "ROLL_State".M[110, 3]) AND (NOT "ROLL_State".M[110, 4]) AND "ROLL_State".M[44, 2]) OR ((NOT "ROLL_State".M[110, 4]) AND "ROLL_State".M[45, 7]) OR "ROLL_State".M[47, 2]);
    "ROLL_State".M[240, 0] := #r;
    // PB10, STEP 5 network 14
    #r := ((NOT "ROLL_IO".Input[119, 7]) AND "ROLL_IO".Input[12, 5] AND "ROLL_IO".Input[12, 7] AND "ROLL_State".M[110, 5] AND "ROLL_State".M[240, 0] AND "ROLL_State".M[35, 2]);
    IF #r THEN "ROLL_State".M[47, 6] := TRUE; END_IF;
    #r := ("ROLL_State".M[32, 2] OR "ROLL_State".M[47, 7]);
    IF #r THEN "ROLL_State".M[47, 6] := FALSE; END_IF;
    // PB10, STEP 5 network 15
    #r := ("ROLL_IO".Input[11, 6] AND "ROLL_IO".Input[119, 7] AND "ROLL_State".M[35, 2] AND "ROLL_State".M[47, 6]);
    IF #r THEN "ROLL_State".M[47, 7] := TRUE; END_IF;
    #r := ("ROLL_State".M[32, 2] OR "ROLL_State".M[48, 0]);
    IF #r THEN "ROLL_State".M[47, 7] := FALSE; END_IF;
    // PB10, STEP 5 network 16
    #r := ((NOT "ROLL_IO".Input[12, 1]) AND "ROLL_IO".Input[12, 5] AND "ROLL_State".M[35, 2] AND "ROLL_State".M[47, 7]);
    IF #r THEN "ROLL_State".M[48, 0] := TRUE; END_IF;
    #r := ("ROLL_State".M[32, 2] OR "ROLL_State".M[48, 1]);
    IF #r THEN "ROLL_State".M[48, 0] := FALSE; END_IF;
    // PB10, STEP 5 network 17
    #r := ("ROLL_IO".Input[12, 1] AND "ROLL_IO".Input[12, 7] AND "ROLL_State".M[35, 2] AND "ROLL_State".M[48, 0]);
    IF #r THEN "ROLL_State".M[48, 1] := TRUE; END_IF;
    #r := ("ROLL_State".M[32, 2] OR "ROLL_State".M[48, 2]);
    IF #r THEN "ROLL_State".M[48, 1] := FALSE; END_IF;
    // PB10, STEP 5 network 18
    #r := ("ROLL_State".M[35, 2] AND "ROLL_State".M[48, 1] AND "ROLL_State".S5Timers[1].Q);
    IF #r THEN "ROLL_State".M[48, 2] := TRUE; END_IF;
    #r := ("ROLL_State".M[32, 2] OR "ROLL_State".M[48, 3]);
    IF #r THEN "ROLL_State".M[48, 2] := FALSE; END_IF;
    // PB10, STEP 5 network 19
    #r := ("ROLL_State".M[35, 2] AND "ROLL_State".M[48, 2]);
    IF #r THEN "ROLL_State".M[48, 3] := TRUE; END_IF;
    #r := ("ROLL_State".M[32, 2] OR "ROLL_State".M[48, 4]);
    IF #r THEN "ROLL_State".M[48, 3] := FALSE; END_IF;
    // PB10, STEP 5 network 20
    #r := ((NOT "ROLL_IO".Input[12, 5]) AND "ROLL_State".M[35, 2] AND "ROLL_State".M[48, 3]);
    IF #r THEN "ROLL_State".M[48, 4] := TRUE; END_IF;
    #r := ("ROLL_State".M[32, 2] OR "ROLL_State".M[48, 5]);
    IF #r THEN "ROLL_State".M[48, 4] := FALSE; END_IF;
    // PB10, STEP 5 network 21
    #r := ("ROLL_IO".Input[12, 5] AND "ROLL_IO".Input[12, 7] AND "ROLL_State".M[35, 2] AND "ROLL_State".M[48, 4]);
    IF #r THEN "ROLL_State".M[48, 5] := TRUE; END_IF;
    #r := ("ROLL_State".M[32, 2] OR "ROLL_State".M[48, 6]);
    IF #r THEN "ROLL_State".M[48, 5] := FALSE; END_IF;
    // PB10, STEP 5 network 22
    #r := ("ROLL_State".M[35, 2] AND "ROLL_State".M[48, 5] AND "ROLL_State".S5Timers[2].Q);
    IF #r THEN "ROLL_State".M[48, 6] := TRUE; END_IF;
    #r := ("ROLL_State".M[32, 2] OR "ROLL_State".M[48, 7] OR "ROLL_State".M[49, 2]);
    IF #r THEN "ROLL_State".M[48, 6] := FALSE; END_IF;
    // PB10, STEP 5 network 23
    #r := ((NOT "ROLL_State".M[110, 6]) AND "ROLL_State".M[35, 2] AND "ROLL_State".M[48, 6]);
    IF #r THEN "ROLL_State".M[48, 7] := TRUE; END_IF;
    #r := ("ROLL_State".M[32, 2] OR "ROLL_State".M[49, 0]);
    IF #r THEN "ROLL_State".M[48, 7] := FALSE; END_IF;
    // PB10, STEP 5 network 24
    #r := ("ROLL_IO".Input[13, 3] AND "ROLL_State".M[35, 2] AND "ROLL_State".M[48, 7] AND "ROLL_State".M[63, 1]);
    IF #r THEN "ROLL_State".M[49, 0] := TRUE; END_IF;
    #r := ("ROLL_State".M[32, 2] OR "ROLL_State".M[50, 6] OR "ROLL_State".M[52, 0]);
    IF #r THEN "ROLL_State".M[49, 0] := FALSE; END_IF;
    // PB10, STEP 5 network 25
    #r := (((NOT "ROLL_State".M[110, 0]) AND (NOT "ROLL_State".M[110, 1]) AND (NOT "ROLL_State".M[110, 2]) AND (NOT "ROLL_State".M[110, 3]) AND (NOT "ROLL_State".M[110, 4]) AND (NOT "ROLL_State".M[110, 5]) AND "ROLL_State".M[40, 1]) OR ((NOT "ROLL_State".M[110, 1]) AND (NOT "ROLL_State".M[110, 2]) AND (NOT "ROLL_State".M[110, 3]) AND (NOT "ROLL_State".M[110, 4]) AND (NOT "ROLL_State".M[110, 5]) AND "ROLL_State".M[41, 2]) OR ((NOT "ROLL_State".M[110, 2]) AND (NOT "ROLL_State".M[110, 3]) AND (NOT "ROLL_State".M[110, 4]) AND (NOT "ROLL_State".M[110, 5]) AND "ROLL_State".M[42, 6]) OR ((NOT "ROLL_State".M[110, 3]) AND (NOT "ROLL_State".M[110, 4]) AND (NOT "ROLL_State".M[110, 5]) AND "ROLL_State".M[44, 2]) OR ((NOT "ROLL_State".M[110, 4]) AND (NOT "ROLL_State".M[110, 5]) AND "ROLL_State".M[45, 7]) OR ((NOT "ROLL_State".M[110, 5]) AND "ROLL_State".M[47, 2]) OR "ROLL_State".M[48, 6]);
    "ROLL_State".M[240, 0] := #r;
    // PB10, STEP 5 network 26
    #r := ((NOT "ROLL_IO".Input[120, 0]) AND "ROLL_IO".Input[12, 5] AND "ROLL_IO".Input[12, 7] AND "ROLL_State".M[110, 6] AND "ROLL_State".M[240, 0] AND "ROLL_State".M[35, 2]);
    IF #r THEN "ROLL_State".M[49, 2] := TRUE; END_IF;
    #r := ("ROLL_State".M[32, 2] OR "ROLL_State".M[49, 3]);
    IF #r THEN "ROLL_State".M[49, 2] := FALSE; END_IF;
    // PB10, STEP 5 network 27
    #r := ("ROLL_IO".Input[11, 6] AND "ROLL_IO".Input[120, 0] AND "ROLL_State".M[35, 2] AND "ROLL_State".M[49, 2]);
    IF #r THEN "ROLL_State".M[49, 3] := TRUE; END_IF;
    #r := ("ROLL_State".M[32, 2] OR "ROLL_State".M[49, 4]);
    IF #r THEN "ROLL_State".M[49, 3] := FALSE; END_IF;
    // PB10, STEP 5 network 28
    #r := ((NOT "ROLL_IO".Input[12, 1]) AND "ROLL_IO".Input[12, 5] AND "ROLL_State".M[35, 2] AND "ROLL_State".M[49, 3]);
    IF #r THEN "ROLL_State".M[49, 4] := TRUE; END_IF;
    #r := ("ROLL_State".M[32, 2] OR "ROLL_State".M[49, 5]);
    IF #r THEN "ROLL_State".M[49, 4] := FALSE; END_IF;
    // PB10, STEP 5 network 29
    #r := ("ROLL_IO".Input[12, 1] AND "ROLL_IO".Input[12, 7] AND "ROLL_State".M[35, 2] AND "ROLL_State".M[49, 4]);
    IF #r THEN "ROLL_State".M[49, 5] := TRUE; END_IF;
    #r := ("ROLL_State".M[32, 2] OR "ROLL_State".M[49, 6]);
    IF #r THEN "ROLL_State".M[49, 5] := FALSE; END_IF;
    // PB10, STEP 5 network 30
    #r := ("ROLL_State".M[35, 2] AND "ROLL_State".M[49, 5] AND "ROLL_State".S5Timers[1].Q);
    IF #r THEN "ROLL_State".M[49, 6] := TRUE; END_IF;
    #r := ("ROLL_State".M[32, 2] OR "ROLL_State".M[49, 7]);
    IF #r THEN "ROLL_State".M[49, 6] := FALSE; END_IF;
    // PB10, STEP 5 network 31
    #r := ("ROLL_State".M[35, 2] AND "ROLL_State".M[49, 6]);
    IF #r THEN "ROLL_State".M[49, 7] := TRUE; END_IF;
    #r := ("ROLL_State".M[32, 2] OR "ROLL_State".M[50, 0]);
    IF #r THEN "ROLL_State".M[49, 7] := FALSE; END_IF;
    // PB10, STEP 5 network 32
    #r := ((NOT "ROLL_IO".Input[12, 5]) AND "ROLL_State".M[35, 2] AND "ROLL_State".M[49, 7]);
    IF #r THEN "ROLL_State".M[50, 0] := TRUE; END_IF;
    #r := ("ROLL_State".M[32, 2] OR "ROLL_State".M[50, 1]);
    IF #r THEN "ROLL_State".M[50, 0] := FALSE; END_IF;
    // PB10, STEP 5 network 33
    #r := ("ROLL_IO".Input[12, 5] AND "ROLL_IO".Input[12, 7] AND "ROLL_State".M[35, 2] AND "ROLL_State".M[50, 0]);
    IF #r THEN "ROLL_State".M[50, 1] := TRUE; END_IF;
    #r := ("ROLL_State".M[32, 2] OR "ROLL_State".M[50, 2]);
    IF #r THEN "ROLL_State".M[50, 1] := FALSE; END_IF;
    // PB10, STEP 5 network 34
    #r := ("ROLL_State".M[35, 2] AND "ROLL_State".M[50, 1] AND "ROLL_State".S5Timers[2].Q);
    IF #r THEN "ROLL_State".M[50, 2] := TRUE; END_IF;
    #r := ("ROLL_State".M[32, 2] OR "ROLL_State".M[50, 3]);
    IF #r THEN "ROLL_State".M[50, 2] := FALSE; END_IF;
    // PB10, STEP 5 network 35
    #r := ("ROLL_State".M[35, 2] AND "ROLL_State".M[50, 2]);
    IF #r THEN "ROLL_State".M[50, 3] := TRUE; END_IF;
    #r := ("ROLL_State".M[32, 2] OR "ROLL_State".M[50, 4]);
    IF #r THEN "ROLL_State".M[50, 3] := FALSE; END_IF;
    // PB10, STEP 5 network 36
    #r := ("ROLL_IO".Input[13, 3] AND "ROLL_State".M[35, 2] AND "ROLL_State".M[50, 3] AND "ROLL_State".M[63, 1]);
    IF #r THEN "ROLL_State".M[50, 4] := TRUE; END_IF;
    #r := ("ROLL_State".M[32, 2] OR "ROLL_State".M[50, 6] OR "ROLL_State".M[52, 0]);
    IF #r THEN "ROLL_State".M[50, 4] := FALSE; END_IF;
    // PB10, STEP 5 network 37
    #r := (((NOT "ROLL_State".M[110, 0]) AND (NOT "ROLL_State".M[110, 1]) AND (NOT "ROLL_State".M[110, 2]) AND (NOT "ROLL_State".M[110, 3]) AND (NOT "ROLL_State".M[110, 4]) AND (NOT "ROLL_State".M[110, 5]) AND (NOT "ROLL_State".M[110, 6]) AND "ROLL_State".M[40, 1]) OR ((NOT "ROLL_State".M[110, 1]) AND (NOT "ROLL_State".M[110, 2]) AND (NOT "ROLL_State".M[110, 3]) AND (NOT "ROLL_State".M[110, 4]) AND (NOT "ROLL_State".M[110, 5]) AND (NOT "ROLL_State".M[110, 6]) AND "ROLL_State".M[41, 4]) OR ((NOT "ROLL_State".M[110, 2]) AND (NOT "ROLL_State".M[110, 3]) AND (NOT "ROLL_State".M[110, 4]) AND (NOT "ROLL_State".M[110, 5]) AND (NOT "ROLL_State".M[110, 6]) AND "ROLL_State".M[43, 0]));
    "ROLL_State".M[240, 0] := #r;
    // PB10, STEP 5 network 38
    #r := (((NOT "ROLL_State".M[110, 3]) AND (NOT "ROLL_State".M[110, 4]) AND (NOT "ROLL_State".M[110, 5]) AND (NOT "ROLL_State".M[110, 6]) AND "ROLL_State".M[44, 4]) OR ((NOT "ROLL_State".M[110, 4]) AND (NOT "ROLL_State".M[110, 5]) AND (NOT "ROLL_State".M[110, 6]) AND "ROLL_State".M[46, 1]) OR ((NOT "ROLL_State".M[110, 5]) AND (NOT "ROLL_State".M[110, 6]) AND "ROLL_State".M[47, 4]) OR ((NOT "ROLL_State".M[110, 6]) AND "ROLL_State".M[49, 0]) OR "ROLL_State".M[50, 4]);
    "ROLL_State".M[240, 1] := #r;
    // PB10, STEP 5 network 39
    #r := ((NOT "ROLL_IO".Input[120, 1]) AND ("ROLL_State".M[240, 0] OR "ROLL_State".M[240, 1]) AND "ROLL_IO".Input[12, 5] AND "ROLL_IO".Input[12, 7] AND "ROLL_State".M[110, 7] AND "ROLL_State".M[35, 2] AND "ROLL_State".M[63, 1]);
    IF #r THEN "ROLL_State".M[50, 6] := TRUE; END_IF;
    #r := ("ROLL_State".M[32, 2] OR "ROLL_State".M[50, 7]);
    IF #r THEN "ROLL_State".M[50, 6] := FALSE; END_IF;
    // PB10, STEP 5 network 40
    #r := ("ROLL_IO".Input[11, 6] AND "ROLL_IO".Input[120, 1] AND "ROLL_State".M[35, 2] AND "ROLL_State".M[50, 6]);
    IF #r THEN "ROLL_State".M[50, 7] := TRUE; END_IF;
    #r := ("ROLL_State".M[32, 2] OR "ROLL_State".M[51, 0]);
    IF #r THEN "ROLL_State".M[50, 7] := FALSE; END_IF;
    // PB10, STEP 5 network 41
    #r := ((NOT "ROLL_IO".Input[12, 1]) AND "ROLL_IO".Input[12, 5] AND "ROLL_State".M[35, 2] AND "ROLL_State".M[50, 7]);
    IF #r THEN "ROLL_State".M[51, 0] := TRUE; END_IF;
    #r := ("ROLL_State".M[32, 2] OR "ROLL_State".M[51, 1]);
    IF #r THEN "ROLL_State".M[51, 0] := FALSE; END_IF;
    // PB10, STEP 5 network 42
    #r := ("ROLL_State".M[35, 2] AND "ROLL_State".M[51, 0] AND "ROLL_State".M[80, 6]);
    IF #r THEN "ROLL_State".M[51, 1] := TRUE; END_IF;
    #r := ("ROLL_State".M[32, 2] OR "ROLL_State".M[51, 2]);
    IF #r THEN "ROLL_State".M[51, 1] := FALSE; END_IF;
    // PB10, STEP 5 network 43
    #r := ("ROLL_State".M[35, 2] AND "ROLL_State".M[51, 1] AND "ROLL_State".S5Timers[1].Q);
    IF #r THEN "ROLL_State".M[51, 2] := TRUE; END_IF;
    #r := ("ROLL_State".M[32, 2] OR "ROLL_State".M[51, 3]);
    IF #r THEN "ROLL_State".M[51, 2] := FALSE; END_IF;
    // PB10, STEP 5 network 44
    #r := ((NOT "ROLL_IO".Input[12, 5]) AND "ROLL_State".M[35, 2] AND "ROLL_State".M[51, 2]);
    IF #r THEN "ROLL_State".M[51, 3] := TRUE; END_IF;
    #r := ("ROLL_State".M[32, 2] OR "ROLL_State".M[51, 4]);
    IF #r THEN "ROLL_State".M[51, 3] := FALSE; END_IF;
    // PB10, STEP 5 network 45
    #r := ("ROLL_IO".Input[12, 5] AND "ROLL_IO".Input[12, 7] AND "ROLL_State".M[35, 2] AND "ROLL_State".M[51, 3]);
    IF #r THEN "ROLL_State".M[51, 4] := TRUE; END_IF;
    #r := ("ROLL_State".M[32, 2] OR "ROLL_State".M[51, 5]);
    IF #r THEN "ROLL_State".M[51, 4] := FALSE; END_IF;
    // PB10, STEP 5 network 46
    #r := ("ROLL_State".M[35, 2] AND "ROLL_State".M[51, 4]);
    IF #r THEN "ROLL_State".M[51, 5] := TRUE; END_IF;
    #r := ("ROLL_State".M[32, 2] OR "ROLL_State".M[51, 6]);
    IF #r THEN "ROLL_State".M[51, 5] := FALSE; END_IF;
    // PB10, STEP 5 network 47
    #r := ("ROLL_IO".Input[13, 3] AND "ROLL_State".M[35, 2] AND "ROLL_State".M[51, 5] AND "ROLL_State".M[63, 1]);
    IF #r THEN "ROLL_State".M[51, 6] := TRUE; END_IF;
    #r := ("ROLL_State".M[32, 2] OR "ROLL_State".M[52, 0]);
    IF #r THEN "ROLL_State".M[51, 6] := FALSE; END_IF;
    // PB10, STEP 5 network 48
    #r := (((NOT "ROLL_State".M[110, 1]) AND (NOT "ROLL_State".M[110, 2]) AND (NOT "ROLL_State".M[110, 3]) AND (NOT "ROLL_State".M[110, 4]) AND (NOT "ROLL_State".M[110, 5]) AND (NOT "ROLL_State".M[110, 6]) AND (NOT "ROLL_State".M[110, 7]) AND "ROLL_State".M[41, 4]) OR ((NOT "ROLL_State".M[110, 2]) AND (NOT "ROLL_State".M[110, 3]) AND (NOT "ROLL_State".M[110, 4]) AND (NOT "ROLL_State".M[110, 5]) AND (NOT "ROLL_State".M[110, 6]) AND (NOT "ROLL_State".M[110, 7]) AND "ROLL_State".M[43, 0]));
    "ROLL_State".M[240, 0] := #r;
    // PB10, STEP 5 network 49
    #r := (((NOT "ROLL_State".M[110, 3]) AND (NOT "ROLL_State".M[110, 4]) AND (NOT "ROLL_State".M[110, 5]) AND (NOT "ROLL_State".M[110, 6]) AND (NOT "ROLL_State".M[110, 7]) AND "ROLL_State".M[44, 4]) OR ((NOT "ROLL_State".M[110, 4]) AND (NOT "ROLL_State".M[110, 5]) AND (NOT "ROLL_State".M[110, 6]) AND (NOT "ROLL_State".M[110, 7]) AND "ROLL_State".M[46, 1]) OR ((NOT "ROLL_State".M[110, 5]) AND (NOT "ROLL_State".M[110, 6]) AND (NOT "ROLL_State".M[110, 7]) AND "ROLL_State".M[47, 4]) OR ((NOT "ROLL_State".M[110, 6]) AND (NOT "ROLL_State".M[110, 7]) AND "ROLL_State".M[49, 0]) OR ((NOT "ROLL_State".M[110, 7]) AND "ROLL_State".M[50, 4]) OR "ROLL_State".M[51, 6]);
    "ROLL_State".M[240, 1] := #r;
    // PB10, STEP 5 network 50
    #r := ((NOT "ROLL_IO".Input[11, 0]) AND ("ROLL_State".M[240, 0] OR "ROLL_State".M[240, 1]) AND "ROLL_IO".Input[12, 5] AND "ROLL_IO".Input[12, 7] AND "ROLL_IO".Input[13, 3] AND "ROLL_State".M[35, 2] AND "ROLL_State".M[63, 1]);
    IF #r THEN "ROLL_State".M[52, 0] := TRUE; END_IF;
    #r := ("ROLL_State".M[32, 2] OR "ROLL_State".M[52, 1]);
    IF #r THEN "ROLL_State".M[52, 0] := FALSE; END_IF;
    // PB10, STEP 5 network 51
    #r := ("ROLL_IO".Input[11, 0] AND "ROLL_IO".Input[11, 6] AND "ROLL_State".M[35, 2] AND "ROLL_State".M[52, 0]);
    IF #r THEN "ROLL_State".M[52, 1] := TRUE; END_IF;
    #r := ("ROLL_State".M[32, 2] OR "ROLL_State".M[52, 2]);
    IF #r THEN "ROLL_State".M[52, 1] := FALSE; END_IF;
    // PB10, STEP 5 network 52
    #r := ((NOT "ROLL_IO".Input[12, 1]) AND (("ROLL_IO".Input[124, 2] AND "ROLL_IO".Input[124, 5]) OR "ROLL_State".M[0, 4]) AND "ROLL_IO".Input[12, 5] AND "ROLL_State".M[35, 2] AND "ROLL_State".M[52, 1]);
    IF #r THEN "ROLL_State".M[52, 2] := TRUE; END_IF;
    #r := ("ROLL_State".M[32, 2] OR "ROLL_State".M[52, 3]);
    IF #r THEN "ROLL_State".M[52, 2] := FALSE; END_IF;
    // PB10, STEP 5 network 53
    #r := ("ROLL_IO".Input[12, 1] AND "ROLL_IO".Input[12, 7] AND "ROLL_State".M[35, 2] AND "ROLL_State".M[52, 2]);
    IF #r THEN "ROLL_State".M[52, 3] := TRUE; END_IF;
    #r := ("ROLL_State".M[32, 2] OR "ROLL_State".M[53, 0] OR "ROLL_State".M[53, 6]);
    IF #r THEN "ROLL_State".M[52, 3] := FALSE; END_IF;
    // PB10, STEP 5 network 54
    #r := ((NOT "ROLL_IO".Output[113, 3]) AND (NOT "ROLL_IO".Input[123, 5]) AND (NOT "ROLL_IO".Input[123, 6]) AND (NOT "ROLL_IO".Input[124, 1]) AND (NOT "ROLL_State".M[70, 3]) AND "ROLL_IO".Output[113, 2] AND "ROLL_IO".Input[124, 2] AND "ROLL_State".M[0, 3] AND "ROLL_State".M[35, 2] AND "ROLL_State".M[52, 3]);
    IF #r THEN "ROLL_State".M[53, 0] := TRUE; END_IF;
    #r := ("ROLL_State".M[32, 2] OR "ROLL_State".M[53, 1]);
    IF #r THEN "ROLL_State".M[53, 0] := FALSE; END_IF;
    // PB10, STEP 5 network 55
    #r := ((NOT "ROLL_IO".Input[124, 2]) AND "ROLL_IO".Input[124, 1] AND "ROLL_State".M[35, 2] AND "ROLL_State".M[53, 0]);
    IF #r THEN "ROLL_State".M[53, 1] := TRUE; END_IF;
    #r := ("ROLL_State".M[32, 2] OR "ROLL_State".M[53, 2]);
    IF #r THEN "ROLL_State".M[53, 1] := FALSE; END_IF;
    // PB10, STEP 5 network 56
    #r := ((NOT "ROLL_IO".Input[124, 4]) AND "ROLL_IO".Input[124, 5] AND "ROLL_State".M[35, 2] AND "ROLL_State".M[53, 1]);
    IF #r THEN "ROLL_State".M[53, 2] := TRUE; END_IF;
    #r := ("ROLL_State".M[32, 2] OR "ROLL_State".M[53, 3]);
    IF #r THEN "ROLL_State".M[53, 2] := FALSE; END_IF;
    // PB10, STEP 5 network 57
    #r := ((NOT "ROLL_IO".Input[124, 5]) AND "ROLL_IO".Input[124, 4] AND "ROLL_State".M[35, 2] AND "ROLL_State".M[53, 2]);
    IF #r THEN "ROLL_State".M[53, 3] := TRUE; END_IF;
    #r := ("ROLL_State".M[32, 2] OR "ROLL_State".M[53, 4]);
    IF #r THEN "ROLL_State".M[53, 3] := FALSE; END_IF;
    // PB10, STEP 5 network 58
    #r := ((NOT "ROLL_State".M[53, 2]) AND "ROLL_State".M[35, 2] AND "ROLL_State".M[53, 3]);
    IF #r THEN "ROLL_State".M[53, 4] := TRUE; END_IF;
    #r := ("ROLL_State".M[32, 2] OR "ROLL_State".M[53, 5]);
    IF #r THEN "ROLL_State".M[53, 4] := FALSE; END_IF;
    // PB10, STEP 5 network 59
    #r := ((NOT "ROLL_IO".Input[123, 5]) AND (NOT "ROLL_IO".Input[123, 6]) AND (NOT "ROLL_State".M[70, 3]) AND "ROLL_State".M[35, 2] AND "ROLL_State".M[53, 4]);
    IF #r THEN "ROLL_State".M[53, 5] := TRUE; END_IF;
    #r := ("ROLL_State".M[32, 2] OR "ROLL_State".M[53, 6]);
    IF #r THEN "ROLL_State".M[53, 5] := FALSE; END_IF;
    // PB10, STEP 5 network 60
    #r := (("ROLL_State".M[52, 3] OR "ROLL_State".M[53, 5]) AND "ROLL_State".M[35, 2]);
    IF #r THEN "ROLL_State".M[53, 6] := TRUE; END_IF;
    #r := ("ROLL_State".M[32, 2] OR "ROLL_State".M[37, 0]);
    IF #r THEN "ROLL_State".M[53, 6] := FALSE; END_IF;
    // PB10, STEP 5 network 61
    RETURN;
END_FUNCTION

